(* PLC project Gaia V5.project, CODESYS CODESYS V3.5 SP22 Patch 2 *)
(* stored: creationDateTime 2026-10-19T15:55:08.3177105, modificationDateTime 2026-10-19T13:52:28.0800332 *)

TYPE DUT_EXC_DOSENSOR : STRUCT
  EXC_OUTPUT_SIGNAL : REAL;  (* [EXC : to other equipment] Dissolved oxygen measure *)
  UPI_INPUT_GLOBAL_LOCAL_FUXA : BOOL;  (* [UPI : functional units to equipment] From UPI_LOCAL_FUXA : global FUXA local active *)
  UPI_INPUT_GLOBAL_LOCAL_HMI : BOOL;  (* From UPI_LOCAL_HMI : global HMI local active *)
  UPI_INPUT_GLOBAL_LOCAL_WEBVISU : BOOL;  (* From UPI_LOCAL_webvisu : global HMI local active *)
END_STRUCT;
END_TYPE

TYPE DUT_IO_DOSENSOR : STRUCT
  INPUT_SIGNAL : DWORD;  (* [INPUT (field to PLC)] Analog input, raw value *)
  INPUT_SENSOR_FAULT : BOOL;  (* Digital input, sensor fault *)
  OUTPUT_CALIBRATION_HIGH : BOOL;  (* [OUTPUT (PLC to field)] Digital output, high calibration *)
  OUTPUT_CALIBRATION_LOW : BOOL;  (* Digital output, low calibration *)
END_STRUCT;
END_TYPE

TYPE DUT_INT_DOSENSOR : STRUCT
  FUXA_LOCAL_REQUEST : BOOL;  (* [Control mode] From FUXA : local request (pulse or maintained) *)
  FUXA_AUTO_REQUEST : BOOL;  (* From FUXA : auto request, releases the individual FUXA local *)
  HMI_LOCAL_REQUEST : BOOL;  (* From HMI : local request (pulse or maintained) *)
  HMI_AUTO_REQUEST : BOOL;  (* From HMI : auto request, releases the individual HMI local *)
  GLOBAL_LOCAL_FUXA : BOOL;  (* From UPI_LOCAL_FUXA : global FUXA local active *)
  GLOBAL_LOCAL_HMI : BOOL;  (* From UPI_LOCAL_HMI : global HMI local active *)
  LOCAL_FUXA_INDIVIDUAL : BOOL;  (* Memory : individual FUXA local, set by local request, reset by auto request *)
  LOCAL_HMI_INDIVIDUAL : BOOL;  (* Memory : individual HMI local, set by local request, reset by auto request *)
  LOCAL_HMI : BOOL;  (* Result : equipment in HMI local (individual or global), unless WEBVISU local is active *)
  LOCAL_FUXA : BOOL;  (* Result : equipment in FUXA local (individual or global), unless WEBVISU or HMI local is active *)
  WEBVISU_LOCAL_REQUEST : BOOL;  (* From WEBVISU : local request (pulse or maintained) *)
  WEBVISU_AUTO_REQUEST : BOOL;  (* From WEBVISU : auto request, releases the individual WEBVISU local *)
  LOCAL_WEBVISU_INDIVIDUAL : BOOL;  (* Memory : individual WEBVISU local, set by local request, reset by auto request *)
  LOCAL_WEBVISU : BOOL;  (* Result : equipment in WEBVISU local (individual or global), has priority *)
  AUTO : BOOL;  (* Result : no local mode, commands come from the functional units (UPI) *)
  SIGNAL_RAW : DWORD;  (* [Inputs] Raw analog input *)
  FAULT : BOOL;  (* Sensor fault (digital input) *)
  CALIB_HIGH_REQUEST : BOOL;  (* High calibration request from the active source *)
  CALIB_LOW_REQUEST : BOOL;  (* Low calibration request from the active source *)
  SIGNAL : REAL;  (* [Results] Scaled measure *)
  CALIB_HIGH : BOOL;  (* High calibration pulse to sensor (1 s) *)
  CALIB_LOW : BOOL;  (* Low calibration pulse to sensor (1 s) *)
  CALIB_DONE : BOOL;  (* Calibration done message (5 s) *)
  GLOBAL_LOCAL_WEBVISU : BOOL;  (* From UPI_LOCAL_WEBVISU : global local request *)
END_STRUCT;
END_TYPE

TYPE DUT_COM_DOSENSOR : STRUCT
  SCADA_INPUT_CALIBRATION_HIGH : BOOL;  (* [SCADA (FUXA) : input (to PLC)] Coil 1 | DO Calibration High *)
  SCADA_INPUT_CALIBRATION_LOW : BOOL;  (* Coil 2 | DO Calibration Low *)
  SCADA_INPUT_LOCAL_REQUEST : BOOL;  (* Coil 8 | DO Sensor Local Request *)
  SCADA_INPUT_AUTO_REQUEST : BOOL;  (* Coil 9 | DO Sensor Auto Request *)
  SCADA_OUTPUT_FAULT : BOOL;  (* [SCADA (FUXA) : output (from PLC)] DI 10001 | Do sensor fault *)
  SCADA_OUTPUT_CALIBRATION_DONE : BOOL;  (* DI 10002 | Do sensor calibration done *)
  SCADA_OUTPUT_LOCAL_FUXA_ACTIVE : BOOL;  (* DI 10013 | DO Sensor Local FUXA Active *)
  SCADA_OUTPUT_LOCAL_HMI_ACTIVE : BOOL;  (* DI 10014 | DO Sensor Local HMI Active *)
  SCADA_OUTPUT_SIGNAL : DUT_Union_Real_Word;  (* IR 89-90 | DO Sensor Signal *)
  HMI_INPUT_CALIBRATION_HIGH : BOOL;  (* [HMI (local panel, FUXA address + 1000) : input (to PLC)] Coil 1001 | DO Calibration High *)
  HMI_INPUT_CALIBRATION_LOW : BOOL;  (* Coil 1002 | DO Calibration Low *)
  HMI_INPUT_LOCAL_REQUEST : BOOL;  (* Coil 1008 | DO Sensor Local Request *)
  HMI_INPUT_AUTO_REQUEST : BOOL;  (* Coil 1009 | DO Sensor Auto Request *)
  HMI_OUTPUT_FAULT : BOOL;  (* [HMI (local panel, FUXA address + 1000) : output (from PLC)] DI 11001 | Do sensor fault *)
  HMI_OUTPUT_CALIBRATION_DONE : BOOL;  (* DI 11002 | Do sensor calibration done *)
  HMI_OUTPUT_LOCAL_ACTIVE : BOOL;  (* DI 11014 | DO Sensor Local Active *)
  HMI_OUTPUT_SIGNAL : DUT_Union_Real_Word;  (* IR 1089-1090 | DO Sensor Signal *)
  WEBVISU_INPUT_CALIBRATION_HIGH : BOOL;  (* DO Calibration High *)
  WEBVISU_INPUT_CALIBRATION_LOW : BOOL;  (* DO Calibration Low *)
  WEBVISU_INPUT_LOCAL_REQUEST : BOOL;  (* DO Sensor Local Request *)
  WEBVISU_INPUT_AUTO_REQUEST : BOOL;  (* DO Sensor Auto Request *)
  WEBVISU_OUTPUT_FAULT : BOOL;  (* Do sensor fault *)
  WEBVISU_OUTPUT_CALIBRATION_DONE : BOOL;  (* Do sensor calibration done *)
  WEBVISU_OUTPUT_LOCAL_ACTIVE : BOOL;  (* DO Sensor Local Active *)
  WEBVISU_OUTPUT_SIGNAL : DUT_Union_Real_Word;  (* DO Sensor Signal *)
  WEBVISU_OUTPUT_LOCAL_FUXA_ACTIVE : BOOL;  (* Effective FUXA local mode (masked by WEBVISU and HMI priority) *)
  WEBVISU_OUTPUT_LOCAL_HMI_ACTIVE : BOOL;  (* Effective HMI local mode (masked by WEBVISU priority) *)
END_STRUCT;
END_TYPE

TYPE DUT_INT_ADM100W : STRUCT
  FUXA_LOCAL_REQUEST : BOOL;  (* [Control mode] From FUXA : local request (pulse or maintained) *)
  FUXA_AUTO_REQUEST : BOOL;  (* From FUXA : auto request, releases the individual FUXA local *)
  HMI_LOCAL_REQUEST : BOOL;  (* From HMI : local request (pulse or maintained) *)
  HMI_AUTO_REQUEST : BOOL;  (* From HMI : auto request, releases the individual HMI local *)
  GLOBAL_LOCAL_FUXA : BOOL;  (* From UPI_LOCAL_FUXA : global FUXA local active *)
  GLOBAL_LOCAL_HMI : BOOL;  (* From UPI_LOCAL_HMI : global HMI local active *)
  LOCAL_FUXA_INDIVIDUAL : BOOL;  (* Memory : individual FUXA local, set by local request, reset by auto request *)
  LOCAL_HMI_INDIVIDUAL : BOOL;  (* Memory : individual HMI local, set by local request, reset by auto request *)
  LOCAL_HMI : BOOL;  (* Result : equipment in HMI local (individual or global), unless WEBVISU local is active *)
  LOCAL_FUXA : BOOL;  (* Result : equipment in FUXA local (individual or global), unless WEBVISU or HMI local is active *)
  AUTO : BOOL;  (* Result : no local mode, commands come from the functional units (UPI) *)
  ALARM_1 : BOOL;  (* [Alarms] Alarm 1 status *)
  ALARM_2 : BOOL;  (* Alarm 2 status *)
  ALARM_3 : BOOL;  (* Alarm 3 status *)
  ALARM_4 : BOOL;  (* Alarm 4 status *)
  ALARM_5 : BOOL;  (* Alarm 5 status *)
  ALARM_6 : BOOL;  (* Alarm 6 status *)
  ALARM_7 : BOOL;  (* Alarm 7 status *)
  ALARM_8 : BOOL;  (* Alarm 8 status *)
  ALARM_9 : BOOL;  (* Alarm 9 status *)
  ALARM_10 : BOOL;  (* Alarm 10 status *)
  FREQUENCY : REAL;  (* [Measures] Frequency | Hz *)
  L1_L2_VOLTAGE : REAL;  (* L1-L2 Voltage | V *)
  L1_N_VOLTAGE : REAL;  (* L1-N Voltage | V *)
  L1_CURRENT : REAL;  (* L1 Current | A *)
  L1_ACTIVE_POWER : REAL;  (* L1 Active Power | W *)
  L1_APPARENT_POWER : REAL;  (* L1 Apparent Power | VA *)
  L1_REACTIVE_POWER : REAL;  (* L1 Reactive Power | W *)
  L1_CURRENT_PHASE_ANGLE : REAL;  (* L1 Current Phase Angle | deg *)
  L1_POWER_FACTOR : REAL;  (* L1 Power Factor | - *)
  L1_VOLTAGE_THD : REAL;  (* L1 Voltage THD | % *)
  L1_CURRENT_THD : REAL;  (* L1 Current THD | % *)
  L1_MAX_LOAD : REAL;  (* L1 Max Load | % of 60 A *)
  L1_L2_VOLTAGE_PHASE_ANGLE : REAL;  (* L1-L2 Voltage Phase Angle | deg *)
  L2_L3_VOLTAGE : REAL;  (* L2-L3 Voltage | V *)
  L2_N_VOLTAGE : REAL;  (* L2-N Voltage | V *)
  L2_CURRENT : REAL;  (* L2 Current | A *)
  L2_ACTIVE_POWER : REAL;  (* L2 Active Power | W *)
  L2_APPARENT_POWER : REAL;  (* L2 Apparent Power | VA *)
  L2_REACTIVE_POWER : REAL;  (* L2 Reactive Power | W *)
  L2_CURRENT_PHASE_ANGLE : REAL;  (* L2 Current Phase Angle | deg *)
  L2_POWER_FACTOR : REAL;  (* L2 Power Factor | - *)
  L2_VOLTAGE_THD : REAL;  (* L2 Voltage THD | % *)
  L2_CURRENT_THD : REAL;  (* L2 Current THD | % *)
  L2_MAX_LOAD : REAL;  (* L2 Max Load | % of 60 A *)
  L1_L3_VOLTAGE_PHASE_ANGLE : REAL;  (* L1-L3 Voltage Phase Angle | deg *)
  L3_L1_VOLTAGE : REAL;  (* L3-L1 Voltage | V *)
  L3_N_VOLTAGE : REAL;  (* L3-N Voltage | V *)
  L3_CURRENT : REAL;  (* L3 Current | A *)
  L3_ACTIVE_POWER : REAL;  (* L3 Active Power | W *)
  L3_APPARENT_POWER : REAL;  (* L3 Apparent Power | VA *)
  L3_REACTIVE_POWER : REAL;  (* L3 Reactive Power | W *)
  L3_CURRENT_PHASE_ANGLE : REAL;  (* L3 Current Phase Angle | deg *)
  L3_POWER_FACTOR : REAL;  (* L3 Power Factor | - *)
  L3_VOLTAGE_THD : REAL;  (* L3 Voltage THD | % *)
  L3_CURRENT_THD : REAL;  (* L3 Current THD | % *)
  L3_MAX_LOAD : REAL;  (* L3 Max Load | % of 60 A *)
  INTERNAL_TEMPERATURE : REAL;  (* Internal Temperature | degC *)
  ACTIVE_ENERGY : REAL;  (* Active Energy | kWh *)
  APPARENT_ENERGY : REAL;  (* Apparent Energy | per ADM100W config *)
  REACTIVE_ENERGY : REAL;  (* Reactive Energy | kWh *)
  TOTAL_ACTIVE_POWER : REAL;  (* Total Active Power | W *)
  TOTAL_APPARENT_POWER : REAL;  (* Total Apparent Power | VA *)
  TOTAL_REACTIVE_POWER : REAL;  (* Total Reactive Power | W *)
  ALL_PHASE_POWER_FACTOR : REAL;  (* All Phase Power Factor | - *)
  WEBVISU_LOCAL_REQUEST : BOOL;  (* From WEBVISU : individual local request *)
  WEBVISU_AUTO_REQUEST : BOOL;  (* From WEBVISU : releases individual WEBVISU local (auto wins) *)
  GLOBAL_LOCAL_WEBVISU : BOOL;  (* From UPI_LOCAL_WEBVISU : global local request *)
  LOCAL_WEBVISU_INDIVIDUAL : BOOL;  (* Memory : individual WEBVISU local request *)
  LOCAL_WEBVISU : BOOL;  (* Effective WEBVISU local : highest source priority *)
END_STRUCT;
END_TYPE

TYPE DUT_COM_UPI_LOCAL_FUXA : STRUCT
  SCADA_INPUT_LOCAL_REQUEST : BOOL;  (* [SCADA (FUXA) : input (to PLC)] Coil 14 | Global Local FUXA Request *)
  SCADA_INPUT_AUTO_REQUEST : BOOL;  (* Coil 15 | Global Auto FUXA Request *)
  SCADA_OUTPUT_LOCAL_ACTIVE : BOOL;  (* [SCADA (FUXA) : output (from PLC)] DI 10019 | Global Local FUXA Active *)
END_STRUCT;
END_TYPE

TYPE DUT_IO_ADM100W : STRUCT
  SPARE : BOOL;  (* Placeholder, structure not used yet *)
END_STRUCT;
END_TYPE

TYPE DUT_COM_ADM100W : STRUCT
  COM_INPUT_IR : ARRAY[0..87] OF WORD;  (* [COM : Modbus RTU, input (equipment to PLC)] Input registers 0..87, 32-bit float, MSW first (ABCD) *)
  COM_INPUT_COILS : ARRAY[0..1] OF BYTE;  (* Coils 0..9 = alarms 1..10 (byte.bit) *)
  SCADA_INPUT_LOCAL_REQUEST : BOOL;  (* [SCADA (FUXA) : input (to PLC)] Coil 12 | ADM100W Local Request *)
  SCADA_INPUT_AUTO_REQUEST : BOOL;  (* Coil 13 | ADM100W Auto Request *)
  SCADA_OUTPUT_ALARM_1_STATUS : BOOL;  (* [SCADA (FUXA) : output (from PLC)] DI 10003 | ADM100W Alarm 1 Status *)
  SCADA_OUTPUT_ALARM_2_STATUS : BOOL;  (* DI 10004 | ADM100W Alarm 2 Status *)
  SCADA_OUTPUT_ALARM_3_STATUS : BOOL;  (* DI 10005 | ADM100W Alarm 3 Status *)
  SCADA_OUTPUT_ALARM_4_STATUS : BOOL;  (* DI 10006 | ADM100W Alarm 4 Status *)
  SCADA_OUTPUT_ALARM_5_STATUS : BOOL;  (* DI 10007 | ADM100W Alarm 5 Status *)
  SCADA_OUTPUT_ALARM_6_STATUS : BOOL;  (* DI 10008 | ADM100W Alarm 6 Status *)
  SCADA_OUTPUT_ALARM_7_STATUS : BOOL;  (* DI 10009 | ADM100W Alarm 7 Status *)
  SCADA_OUTPUT_ALARM_8_STATUS : BOOL;  (* DI 10010 | ADM100W Alarm 8 Status *)
  SCADA_OUTPUT_ALARM_9_STATUS : BOOL;  (* DI 10011 | ADM100W Alarm 9 Status *)
  SCADA_OUTPUT_ALARM_10_STATUS : BOOL;  (* DI 10012 | ADM100W Alarm 10 Status *)
  SCADA_OUTPUT_LOCAL_FUXA_ACTIVE : BOOL;  (* DI 10017 | ADM100W Local FUXA Active *)
  SCADA_OUTPUT_LOCAL_HMI_ACTIVE : BOOL;  (* DI 10018 | ADM100W Local HMI Active *)
  SCADA_OUTPUT_FREQUENCY : DUT_Union_Real_Word;  (* IR 1-2 | ADM100W Frequency | Hz *)
  SCADA_OUTPUT_L1_L2_VOLTAGE : DUT_Union_Real_Word;  (* IR 3-4 | ADM100W L1-L2 Voltage | V *)
  SCADA_OUTPUT_L1_N_VOLTAGE : DUT_Union_Real_Word;  (* IR 5-6 | ADM100W L1-N Voltage | V *)
  SCADA_OUTPUT_L1_CURRENT : DUT_Union_Real_Word;  (* IR 7-8 | ADM100W L1 Current | A *)
  SCADA_OUTPUT_L1_ACTIVE_POWER : DUT_Union_Real_Word;  (* IR 9-10 | ADM100W L1 Active Power *)
  SCADA_OUTPUT_L1_APPARENT_POWER : DUT_Union_Real_Word;  (* IR 11-12 | ADM100W L1 Apparent Power *)
  SCADA_OUTPUT_L1_REACTIVE_POWER : DUT_Union_Real_Word;  (* IR 13-14 | ADM100W L1 Reactive Power *)
  SCADA_OUTPUT_L1_CURRENT_PHASE_ANGLE : DUT_Union_Real_Word;  (* IR 15-16 | ADM100W L1 Current Phase Angle | deg *)
  SCADA_OUTPUT_L1_POWER_FACTOR : DUT_Union_Real_Word;  (* IR 17-18 | ADM100W L1 Power Factor *)
  SCADA_OUTPUT_L1_VOLTAGE_THD : DUT_Union_Real_Word;  (* IR 19-20 | ADM100W L1 Voltage THD | % *)
  SCADA_OUTPUT_L1_CURRENT_THD : DUT_Union_Real_Word;  (* IR 21-22 | ADM100W L1 Current THD | % *)
  SCADA_OUTPUT_L1_MAX_LOAD : DUT_Union_Real_Word;  (* IR 23-24 | ADM100W L1 Max Load *)
  SCADA_OUTPUT_L1_L2_VOLTAGE_PHASE_ANGLE : DUT_Union_Real_Word;  (* IR 25-26 | ADM100W L1-L2 Voltage Phase Angle | deg *)
  SCADA_OUTPUT_L2_L3_VOLTAGE : DUT_Union_Real_Word;  (* IR 27-28 | ADM100W L2-L3 Voltage | V *)
  SCADA_OUTPUT_L2_N_VOLTAGE : DUT_Union_Real_Word;  (* IR 29-30 | ADM100W L2-N Voltage | V *)
  SCADA_OUTPUT_L2_CURRENT : DUT_Union_Real_Word;  (* IR 31-32 | ADM100W L2 Current | A *)
  SCADA_OUTPUT_L2_ACTIVE_POWER : DUT_Union_Real_Word;  (* IR 33-34 | ADM100W L2 Active Power *)
  SCADA_OUTPUT_L2_APPARENT_POWER : DUT_Union_Real_Word;  (* IR 35-36 | ADM100W L2 Apparent Power *)
  SCADA_OUTPUT_L2_REACTIVE_POWER : DUT_Union_Real_Word;  (* IR 37-38 | ADM100W L2 Reactive Power *)
  SCADA_OUTPUT_L2_CURRENT_PHASE_ANGLE : DUT_Union_Real_Word;  (* IR 39-40 | ADM100W L2 Current Phase Angle | deg *)
  SCADA_OUTPUT_L2_POWER_FACTOR : DUT_Union_Real_Word;  (* IR 41-42 | ADM100W L2 Power Factor *)
  SCADA_OUTPUT_L2_VOLTAGE_THD : DUT_Union_Real_Word;  (* IR 43-44 | ADM100W L2 Voltage THD | % *)
  SCADA_OUTPUT_L2_CURRENT_THD : DUT_Union_Real_Word;  (* IR 45-46 | ADM100W L2 Current THD | % *)
  SCADA_OUTPUT_L2_MAX_LOAD : DUT_Union_Real_Word;  (* IR 47-48 | ADM100W L2 Max Load *)
  SCADA_OUTPUT_L1_L3_VOLTAGE_PHASE_ANGLE : DUT_Union_Real_Word;  (* IR 49-50 | ADM100W L1-L3 Voltage Phase Angle | deg *)
  SCADA_OUTPUT_L3_L1_VOLTAGE : DUT_Union_Real_Word;  (* IR 51-52 | ADM100W L3-L1 Voltage | V *)
  SCADA_OUTPUT_L3_N_VOLTAGE : DUT_Union_Real_Word;  (* IR 53-54 | ADM100W L3-N Voltage | V *)
  SCADA_OUTPUT_L3_CURRENT : DUT_Union_Real_Word;  (* IR 55-56 | ADM100W L3 Current | A *)
  SCADA_OUTPUT_L3_ACTIVE_POWER : DUT_Union_Real_Word;  (* IR 57-58 | ADM100W L3 Active Power *)
  SCADA_OUTPUT_L3_APPARENT_POWER : DUT_Union_Real_Word;  (* IR 59-60 | ADM100W L3 Apparent Power *)
  SCADA_OUTPUT_L3_REACTIVE_POWER : DUT_Union_Real_Word;  (* IR 61-62 | ADM100W L3 Reactive Power *)
  SCADA_OUTPUT_L3_CURRENT_PHASE_ANGLE : DUT_Union_Real_Word;  (* IR 63-64 | ADM100W L3 Current Phase Angle | deg *)
  SCADA_OUTPUT_L3_POWER_FACTOR : DUT_Union_Real_Word;  (* IR 65-66 | ADM100W L3 Power Factor *)
  SCADA_OUTPUT_L3_VOLTAGE_THD : DUT_Union_Real_Word;  (* IR 67-68 | ADM100W L3 Voltage THD | % *)
  SCADA_OUTPUT_L3_CURRENT_THD : DUT_Union_Real_Word;  (* IR 69-70 | ADM100W L3 Current THD | % *)
  SCADA_OUTPUT_L3_MAX_LOAD : DUT_Union_Real_Word;  (* IR 71-72 | ADM100W L3 Max Load *)
  SCADA_OUTPUT_INTERNAL_TEMPERATURE : DUT_Union_Real_Word;  (* IR 73-74 | ADM100W Internal Temperature *)
  SCADA_OUTPUT_ACTIVE_ENERGY : DUT_Union_Real_Word;  (* IR 75-76 | ADM100W Active Energy *)
  SCADA_OUTPUT_APPARENT_ENERGY : DUT_Union_Real_Word;  (* IR 77-78 | ADM100W Apparent Energy *)
  SCADA_OUTPUT_REACTIVE_ENERGY : DUT_Union_Real_Word;  (* IR 79-80 | ADM100W Reactive Energy *)
  SCADA_OUTPUT_TOTAL_ACTIVE_POWER : DUT_Union_Real_Word;  (* IR 81-82 | ADM100W Total Active Power *)
  SCADA_OUTPUT_TOTAL_APPARENT_POWER : DUT_Union_Real_Word;  (* IR 83-84 | ADM100W Total Apparent Power *)
  SCADA_OUTPUT_TOTAL_REACTIVE_POWER : DUT_Union_Real_Word;  (* IR 85-86 | ADM100W Total Reactive Power *)
  SCADA_OUTPUT_ALL_PHASE_POWER_FACTOR : DUT_Union_Real_Word;  (* IR 87-88 | ADM100W All Phase Power Factor *)
  HMI_INPUT_LOCAL_REQUEST : BOOL;  (* [HMI (local panel, FUXA address + 1000) : input (to PLC)] Coil 1012 | ADM100W Local Request *)
  HMI_INPUT_AUTO_REQUEST : BOOL;  (* Coil 1013 | ADM100W Auto Request *)
  HMI_OUTPUT_ALARM_1_STATUS : BOOL;  (* [HMI (local panel, FUXA address + 1000) : output (from PLC)] DI 11003 | ADM100W Alarm 1 Status *)
  HMI_OUTPUT_ALARM_2_STATUS : BOOL;  (* DI 11004 | ADM100W Alarm 2 Status *)
  HMI_OUTPUT_ALARM_3_STATUS : BOOL;  (* DI 11005 | ADM100W Alarm 3 Status *)
  HMI_OUTPUT_ALARM_4_STATUS : BOOL;  (* DI 11006 | ADM100W Alarm 4 Status *)
  HMI_OUTPUT_ALARM_5_STATUS : BOOL;  (* DI 11007 | ADM100W Alarm 5 Status *)
  HMI_OUTPUT_ALARM_6_STATUS : BOOL;  (* DI 11008 | ADM100W Alarm 6 Status *)
  HMI_OUTPUT_ALARM_7_STATUS : BOOL;  (* DI 11009 | ADM100W Alarm 7 Status *)
  HMI_OUTPUT_ALARM_8_STATUS : BOOL;  (* DI 11010 | ADM100W Alarm 8 Status *)
  HMI_OUTPUT_ALARM_9_STATUS : BOOL;  (* DI 11011 | ADM100W Alarm 9 Status *)
  HMI_OUTPUT_ALARM_10_STATUS : BOOL;  (* DI 11012 | ADM100W Alarm 10 Status *)
  HMI_OUTPUT_LOCAL_ACTIVE : BOOL;  (* DI 11018 | ADM100W Local Active *)
  HMI_OUTPUT_FREQUENCY : DUT_Union_Real_Word;  (* IR 1001-1002 | ADM100W Frequency | Hz *)
  HMI_OUTPUT_L1_L2_VOLTAGE : DUT_Union_Real_Word;  (* IR 1003-1004 | ADM100W L1-L2 Voltage | V *)
  HMI_OUTPUT_L1_N_VOLTAGE : DUT_Union_Real_Word;  (* IR 1005-1006 | ADM100W L1-N Voltage | V *)
  HMI_OUTPUT_L1_CURRENT : DUT_Union_Real_Word;  (* IR 1007-1008 | ADM100W L1 Current | A *)
  HMI_OUTPUT_L1_ACTIVE_POWER : DUT_Union_Real_Word;  (* IR 1009-1010 | ADM100W L1 Active Power *)
  HMI_OUTPUT_L1_APPARENT_POWER : DUT_Union_Real_Word;  (* IR 1011-1012 | ADM100W L1 Apparent Power *)
  HMI_OUTPUT_L1_REACTIVE_POWER : DUT_Union_Real_Word;  (* IR 1013-1014 | ADM100W L1 Reactive Power *)
  HMI_OUTPUT_L1_CURRENT_PHASE_ANGLE : DUT_Union_Real_Word;  (* IR 1015-1016 | ADM100W L1 Current Phase Angle | deg *)
  HMI_OUTPUT_L1_POWER_FACTOR : DUT_Union_Real_Word;  (* IR 1017-1018 | ADM100W L1 Power Factor *)
  HMI_OUTPUT_L1_VOLTAGE_THD : DUT_Union_Real_Word;  (* IR 1019-1020 | ADM100W L1 Voltage THD | % *)
  HMI_OUTPUT_L1_CURRENT_THD : DUT_Union_Real_Word;  (* IR 1021-1022 | ADM100W L1 Current THD | % *)
  HMI_OUTPUT_L1_MAX_LOAD : DUT_Union_Real_Word;  (* IR 1023-1024 | ADM100W L1 Max Load *)
  HMI_OUTPUT_L1_L2_VOLTAGE_PHASE_ANGLE : DUT_Union_Real_Word;  (* IR 1025-1026 | ADM100W L1-L2 Voltage Phase Angle | deg *)
  HMI_OUTPUT_L2_L3_VOLTAGE : DUT_Union_Real_Word;  (* IR 1027-1028 | ADM100W L2-L3 Voltage | V *)
  HMI_OUTPUT_L2_N_VOLTAGE : DUT_Union_Real_Word;  (* IR 1029-1030 | ADM100W L2-N Voltage | V *)
  HMI_OUTPUT_L2_CURRENT : DUT_Union_Real_Word;  (* IR 1031-1032 | ADM100W L2 Current | A *)
  HMI_OUTPUT_L2_ACTIVE_POWER : DUT_Union_Real_Word;  (* IR 1033-1034 | ADM100W L2 Active Power *)
  HMI_OUTPUT_L2_APPARENT_POWER : DUT_Union_Real_Word;  (* IR 1035-1036 | ADM100W L2 Apparent Power *)
  HMI_OUTPUT_L2_REACTIVE_POWER : DUT_Union_Real_Word;  (* IR 1037-1038 | ADM100W L2 Reactive Power *)
  HMI_OUTPUT_L2_CURRENT_PHASE_ANGLE : DUT_Union_Real_Word;  (* IR 1039-1040 | ADM100W L2 Current Phase Angle | deg *)
  HMI_OUTPUT_L2_POWER_FACTOR : DUT_Union_Real_Word;  (* IR 1041-1042 | ADM100W L2 Power Factor *)
  HMI_OUTPUT_L2_VOLTAGE_THD : DUT_Union_Real_Word;  (* IR 1043-1044 | ADM100W L2 Voltage THD | % *)
  HMI_OUTPUT_L2_CURRENT_THD : DUT_Union_Real_Word;  (* IR 1045-1046 | ADM100W L2 Current THD | % *)
  HMI_OUTPUT_L2_MAX_LOAD : DUT_Union_Real_Word;  (* IR 1047-1048 | ADM100W L2 Max Load *)
  HMI_OUTPUT_L1_L3_VOLTAGE_PHASE_ANGLE : DUT_Union_Real_Word;  (* IR 1049-1050 | ADM100W L1-L3 Voltage Phase Angle | deg *)
  HMI_OUTPUT_L3_L1_VOLTAGE : DUT_Union_Real_Word;  (* IR 1051-1052 | ADM100W L3-L1 Voltage | V *)
  HMI_OUTPUT_L3_N_VOLTAGE : DUT_Union_Real_Word;  (* IR 1053-1054 | ADM100W L3-N Voltage | V *)
  HMI_OUTPUT_L3_CURRENT : DUT_Union_Real_Word;  (* IR 1055-1056 | ADM100W L3 Current | A *)
  HMI_OUTPUT_L3_ACTIVE_POWER : DUT_Union_Real_Word;  (* IR 1057-1058 | ADM100W L3 Active Power *)
  HMI_OUTPUT_L3_APPARENT_POWER : DUT_Union_Real_Word;  (* IR 1059-1060 | ADM100W L3 Apparent Power *)
  HMI_OUTPUT_L3_REACTIVE_POWER : DUT_Union_Real_Word;  (* IR 1061-1062 | ADM100W L3 Reactive Power *)
  HMI_OUTPUT_L3_CURRENT_PHASE_ANGLE : DUT_Union_Real_Word;  (* IR 1063-1064 | ADM100W L3 Current Phase Angle | deg *)
  HMI_OUTPUT_L3_POWER_FACTOR : DUT_Union_Real_Word;  (* IR 1065-1066 | ADM100W L3 Power Factor *)
  HMI_OUTPUT_L3_VOLTAGE_THD : DUT_Union_Real_Word;  (* IR 1067-1068 | ADM100W L3 Voltage THD | % *)
  HMI_OUTPUT_L3_CURRENT_THD : DUT_Union_Real_Word;  (* IR 1069-1070 | ADM100W L3 Current THD | % *)
  HMI_OUTPUT_L3_MAX_LOAD : DUT_Union_Real_Word;  (* IR 1071-1072 | ADM100W L3 Max Load *)
  HMI_OUTPUT_INTERNAL_TEMPERATURE : DUT_Union_Real_Word;  (* IR 1073-1074 | ADM100W Internal Temperature *)
  HMI_OUTPUT_ACTIVE_ENERGY : DUT_Union_Real_Word;  (* IR 1075-1076 | ADM100W Active Energy *)
  HMI_OUTPUT_APPARENT_ENERGY : DUT_Union_Real_Word;  (* IR 1077-1078 | ADM100W Apparent Energy *)
  HMI_OUTPUT_REACTIVE_ENERGY : DUT_Union_Real_Word;  (* IR 1079-1080 | ADM100W Reactive Energy *)
  HMI_OUTPUT_TOTAL_ACTIVE_POWER : DUT_Union_Real_Word;  (* IR 1081-1082 | ADM100W Total Active Power *)
  HMI_OUTPUT_TOTAL_APPARENT_POWER : DUT_Union_Real_Word;  (* IR 1083-1084 | ADM100W Total Apparent Power *)
  HMI_OUTPUT_TOTAL_REACTIVE_POWER : DUT_Union_Real_Word;  (* IR 1085-1086 | ADM100W Total Reactive Power *)
  HMI_OUTPUT_ALL_PHASE_POWER_FACTOR : DUT_Union_Real_Word;  (* IR 1087-1088 | ADM100W All Phase Power Factor *)
  WEBVISU_INPUT_LOCAL_REQUEST : BOOL;  (* [WEBVISU : direct IEC variable] ADM100W Local Request *)
  WEBVISU_INPUT_AUTO_REQUEST : BOOL;  (* [WEBVISU : direct IEC variable] ADM100W Auto Request *)
  WEBVISU_OUTPUT_ALARM_1_STATUS : BOOL;  (* [WEBVISU : direct IEC variable] ADM100W Alarm 1 Status *)
  WEBVISU_OUTPUT_ALARM_2_STATUS : BOOL;  (* [WEBVISU : direct IEC variable] ADM100W Alarm 2 Status *)
  WEBVISU_OUTPUT_ALARM_3_STATUS : BOOL;  (* [WEBVISU : direct IEC variable] ADM100W Alarm 3 Status *)
  WEBVISU_OUTPUT_ALARM_4_STATUS : BOOL;  (* [WEBVISU : direct IEC variable] ADM100W Alarm 4 Status *)
  WEBVISU_OUTPUT_ALARM_5_STATUS : BOOL;  (* [WEBVISU : direct IEC variable] ADM100W Alarm 5 Status *)
  WEBVISU_OUTPUT_ALARM_6_STATUS : BOOL;  (* [WEBVISU : direct IEC variable] ADM100W Alarm 6 Status *)
  WEBVISU_OUTPUT_ALARM_7_STATUS : BOOL;  (* [WEBVISU : direct IEC variable] ADM100W Alarm 7 Status *)
  WEBVISU_OUTPUT_ALARM_8_STATUS : BOOL;  (* [WEBVISU : direct IEC variable] ADM100W Alarm 8 Status *)
  WEBVISU_OUTPUT_ALARM_9_STATUS : BOOL;  (* [WEBVISU : direct IEC variable] ADM100W Alarm 9 Status *)
  WEBVISU_OUTPUT_ALARM_10_STATUS : BOOL;  (* [WEBVISU : direct IEC variable] ADM100W Alarm 10 Status *)
  WEBVISU_OUTPUT_LOCAL_ACTIVE : BOOL;  (* [WEBVISU : direct IEC variable] ADM100W Local Active *)
  WEBVISU_OUTPUT_FREQUENCY : DUT_Union_Real_Word;  (* [WEBVISU : direct IEC variable] ADM100W Frequency | Hz *)
  WEBVISU_OUTPUT_L1_L2_VOLTAGE : DUT_Union_Real_Word;  (* [WEBVISU : direct IEC variable] ADM100W L1-L2 Voltage | V *)
  WEBVISU_OUTPUT_L1_N_VOLTAGE : DUT_Union_Real_Word;  (* [WEBVISU : direct IEC variable] ADM100W L1-N Voltage | V *)
  WEBVISU_OUTPUT_L1_CURRENT : DUT_Union_Real_Word;  (* [WEBVISU : direct IEC variable] ADM100W L1 Current | A *)
  WEBVISU_OUTPUT_L1_ACTIVE_POWER : DUT_Union_Real_Word;  (* [WEBVISU : direct IEC variable] ADM100W L1 Active Power *)
  WEBVISU_OUTPUT_L1_APPARENT_POWER : DUT_Union_Real_Word;  (* [WEBVISU : direct IEC variable] ADM100W L1 Apparent Power *)
  WEBVISU_OUTPUT_L1_REACTIVE_POWER : DUT_Union_Real_Word;  (* [WEBVISU : direct IEC variable] ADM100W L1 Reactive Power *)
  WEBVISU_OUTPUT_L1_CURRENT_PHASE_ANGLE : DUT_Union_Real_Word;  (* [WEBVISU : direct IEC variable] ADM100W L1 Current Phase Angle | deg *)
  WEBVISU_OUTPUT_L1_POWER_FACTOR : DUT_Union_Real_Word;  (* [WEBVISU : direct IEC variable] ADM100W L1 Power Factor *)
  WEBVISU_OUTPUT_L1_VOLTAGE_THD : DUT_Union_Real_Word;  (* [WEBVISU : direct IEC variable] ADM100W L1 Voltage THD | % *)
  WEBVISU_OUTPUT_L1_CURRENT_THD : DUT_Union_Real_Word;  (* [WEBVISU : direct IEC variable] ADM100W L1 Current THD | % *)
  WEBVISU_OUTPUT_L1_MAX_LOAD : DUT_Union_Real_Word;  (* [WEBVISU : direct IEC variable] ADM100W L1 Max Load *)
  WEBVISU_OUTPUT_L1_L2_VOLTAGE_PHASE_ANGLE : DUT_Union_Real_Word;  (* [WEBVISU : direct IEC variable] ADM100W L1-L2 Voltage Phase Angle | deg *)
  WEBVISU_OUTPUT_L2_L3_VOLTAGE : DUT_Union_Real_Word;  (* [WEBVISU : direct IEC variable] ADM100W L2-L3 Voltage | V *)
  WEBVISU_OUTPUT_L2_N_VOLTAGE : DUT_Union_Real_Word;  (* [WEBVISU : direct IEC variable] ADM100W L2-N Voltage | V *)
  WEBVISU_OUTPUT_L2_CURRENT : DUT_Union_Real_Word;  (* [WEBVISU : direct IEC variable] ADM100W L2 Current | A *)
  WEBVISU_OUTPUT_L2_ACTIVE_POWER : DUT_Union_Real_Word;  (* [WEBVISU : direct IEC variable] ADM100W L2 Active Power *)
  WEBVISU_OUTPUT_L2_APPARENT_POWER : DUT_Union_Real_Word;  (* [WEBVISU : direct IEC variable] ADM100W L2 Apparent Power *)
  WEBVISU_OUTPUT_L2_REACTIVE_POWER : DUT_Union_Real_Word;  (* [WEBVISU : direct IEC variable] ADM100W L2 Reactive Power *)
  WEBVISU_OUTPUT_L2_CURRENT_PHASE_ANGLE : DUT_Union_Real_Word;  (* [WEBVISU : direct IEC variable] ADM100W L2 Current Phase Angle | deg *)
  WEBVISU_OUTPUT_L2_POWER_FACTOR : DUT_Union_Real_Word;  (* [WEBVISU : direct IEC variable] ADM100W L2 Power Factor *)
  WEBVISU_OUTPUT_L2_VOLTAGE_THD : DUT_Union_Real_Word;  (* [WEBVISU : direct IEC variable] ADM100W L2 Voltage THD | % *)
  WEBVISU_OUTPUT_L2_CURRENT_THD : DUT_Union_Real_Word;  (* [WEBVISU : direct IEC variable] ADM100W L2 Current THD | % *)
  WEBVISU_OUTPUT_L2_MAX_LOAD : DUT_Union_Real_Word;  (* [WEBVISU : direct IEC variable] ADM100W L2 Max Load *)
  WEBVISU_OUTPUT_L1_L3_VOLTAGE_PHASE_ANGLE : DUT_Union_Real_Word;  (* [WEBVISU : direct IEC variable] ADM100W L1-L3 Voltage Phase Angle | deg *)
  WEBVISU_OUTPUT_L3_L1_VOLTAGE : DUT_Union_Real_Word;  (* [WEBVISU : direct IEC variable] ADM100W L3-L1 Voltage | V *)
  WEBVISU_OUTPUT_L3_N_VOLTAGE : DUT_Union_Real_Word;  (* [WEBVISU : direct IEC variable] ADM100W L3-N Voltage | V *)
  WEBVISU_OUTPUT_L3_CURRENT : DUT_Union_Real_Word;  (* [WEBVISU : direct IEC variable] ADM100W L3 Current | A *)
  WEBVISU_OUTPUT_L3_ACTIVE_POWER : DUT_Union_Real_Word;  (* [WEBVISU : direct IEC variable] ADM100W L3 Active Power *)
  WEBVISU_OUTPUT_L3_APPARENT_POWER : DUT_Union_Real_Word;  (* [WEBVISU : direct IEC variable] ADM100W L3 Apparent Power *)
  WEBVISU_OUTPUT_L3_REACTIVE_POWER : DUT_Union_Real_Word;  (* [WEBVISU : direct IEC variable] ADM100W L3 Reactive Power *)
  WEBVISU_OUTPUT_L3_CURRENT_PHASE_ANGLE : DUT_Union_Real_Word;  (* [WEBVISU : direct IEC variable] ADM100W L3 Current Phase Angle | deg *)
  WEBVISU_OUTPUT_L3_POWER_FACTOR : DUT_Union_Real_Word;  (* [WEBVISU : direct IEC variable] ADM100W L3 Power Factor *)
  WEBVISU_OUTPUT_L3_VOLTAGE_THD : DUT_Union_Real_Word;  (* [WEBVISU : direct IEC variable] ADM100W L3 Voltage THD | % *)
  WEBVISU_OUTPUT_L3_CURRENT_THD : DUT_Union_Real_Word;  (* [WEBVISU : direct IEC variable] ADM100W L3 Current THD | % *)
  WEBVISU_OUTPUT_L3_MAX_LOAD : DUT_Union_Real_Word;  (* [WEBVISU : direct IEC variable] ADM100W L3 Max Load *)
  WEBVISU_OUTPUT_INTERNAL_TEMPERATURE : DUT_Union_Real_Word;  (* [WEBVISU : direct IEC variable] ADM100W Internal Temperature *)
  WEBVISU_OUTPUT_ACTIVE_ENERGY : DUT_Union_Real_Word;  (* [WEBVISU : direct IEC variable] ADM100W Active Energy *)
  WEBVISU_OUTPUT_APPARENT_ENERGY : DUT_Union_Real_Word;  (* [WEBVISU : direct IEC variable] ADM100W Apparent Energy *)
  WEBVISU_OUTPUT_REACTIVE_ENERGY : DUT_Union_Real_Word;  (* [WEBVISU : direct IEC variable] ADM100W Reactive Energy *)
  WEBVISU_OUTPUT_TOTAL_ACTIVE_POWER : DUT_Union_Real_Word;  (* [WEBVISU : direct IEC variable] ADM100W Total Active Power *)
  WEBVISU_OUTPUT_TOTAL_APPARENT_POWER : DUT_Union_Real_Word;  (* [WEBVISU : direct IEC variable] ADM100W Total Apparent Power *)
  WEBVISU_OUTPUT_TOTAL_REACTIVE_POWER : DUT_Union_Real_Word;  (* [WEBVISU : direct IEC variable] ADM100W Total Reactive Power *)
  WEBVISU_OUTPUT_ALL_PHASE_POWER_FACTOR : DUT_Union_Real_Word;  (* [WEBVISU : direct IEC variable] ADM100W All Phase Power Factor *)
  WEBVISU_OUTPUT_LOCAL_FUXA_ACTIVE : BOOL;  (* Effective FUXA local mode (masked by WEBVISU and HMI priority) *)
  WEBVISU_OUTPUT_LOCAL_HMI_ACTIVE : BOOL;  (* Effective HMI local mode (masked by WEBVISU priority) *)
END_STRUCT;
END_TYPE

TYPE DUT_EXC_ADM100W : STRUCT
  EXC_OUTPUT_FREQUENCY : REAL;  (* [EXC : to other equipment] Hz *)
  EXC_OUTPUT_L1_N_VOLTAGE : REAL;  (* V *)
  EXC_OUTPUT_L1_CURRENT : REAL;  (* A *)
  EXC_OUTPUT_L1_ACTIVE_POWER : REAL;  (* W *)
  EXC_OUTPUT_L1_APPARENT_POWER : REAL;  (* VA *)
  EXC_OUTPUT_L1_REACTIVE_POWER : REAL;  (* VAr *)
  EXC_OUTPUT_L1_POWER_FACTOR : REAL;  (* - *)
  EXC_OUTPUT_L1_VOLTAGE_THD : REAL;  (* % *)
  EXC_OUTPUT_L1_CURRENT_THD : REAL;  (* % *)
  EXC_OUTPUT_L1_MAX_LOAD : REAL;  (* % of 60 A *)
  EXC_OUTPUT_INTERNAL_TEMPERATURE : REAL;  (* degC *)
  EXC_OUTPUT_ACTIVE_ENERGY : REAL;  (* kWh *)
  EXC_OUTPUT_DATA_VALID : BOOL;  (* FALSE = values not usable. Not managed yet (no Modbus diagnostic) *)
  UPI_INPUT_GLOBAL_LOCAL_FUXA : BOOL;  (* [UPI : functional units to equipment] From UPI_LOCAL_FUXA : global FUXA local active *)
  UPI_INPUT_GLOBAL_LOCAL_HMI : BOOL;  (* From UPI_LOCAL_HMI : global HMI local active *)
  UPI_INPUT_GLOBAL_LOCAL_WEBVISU : BOOL;  (* From UPI_LOCAL_WEBVISU : global WEBVISU local active *)
END_STRUCT;
END_TYPE

TYPE DUT_COM_DIP1500 : STRUCT
  COM_INPUT_IR : ARRAY[0..4] OF WORD;  (* [COM : Modbus RTU, input (equipment to PLC)] Input registers 0x3001..0x3005 *)
  COM_INPUT_HR_COUNTERS : ARRAY[0..3] OF WORD;  (* Holding registers 0x4007..0x400A (read) *)
  COM_OUTPUT_COILS : ARRAY[0..3] OF BOOL;  (* [COM : Modbus RTU, output (PLC to equipment)] Coils 0x0001..0x0004 *)
  COM_OUTPUT_HR_CMD : ARRAY[0..5] OF WORD;  (* Holding registers 0x4001..0x4006 (write) *)
  COM_OUTPUT_HR_CONFIG : ARRAY[0..6] OF WORD;  (* Holding registers 0x400B..0x4011 (write) *)
  COM_OUTPUT_CMD_TRIGGER : BOOL;  (* Rising edge trigger of the command write channel(s), mapped in the Modbus slave I/O mapping *)
  COM_OUTPUT_CONFIG_TRIGGER : BOOL;  (* Rising edge trigger of the configuration write channel, mapped in the Modbus slave I/O mapping *)
  SCADA_INPUT_MOTOR_START_STOP : BOOL;  (* [SCADA (FUXA) : input (to PLC)] Coil 3 | DIP1500 Motor Start Stop *)
  SCADA_INPUT_MOTOR_DIRECTION : BOOL;  (* Coil 4 | DIP1500 Motor Direction *)
  SCADA_INPUT_FLASH_SAVE : BOOL;  (* Coil 5 | DIP1500 Flash Save *)
  SCADA_INPUT_OPERATION_MODE : BOOL;  (* Coil 6 | DIP1500 Operation Mode *)
  SCADA_INPUT_PARAM_WRITE_ENABLE : BOOL;  (* Coil 7 | DIP1500 Parameter Write Enable *)
  SCADA_INPUT_LOCAL_REQUEST : BOOL;  (* Coil 10 | DIP1500 Local Request *)
  SCADA_INPUT_AUTO_REQUEST : BOOL;  (* Coil 11 | DIP1500 Auto Request *)
  SCADA_INPUT_FOOT_SWITCH_INPUT_MODE : WORD;  (* HR 9 | DIP1500 Foot Switch Input Mode *)
  SCADA_INPUT_LIQUID_LEVEL_INPUT_MODE : WORD;  (* HR 10 | DIP1500 Liquid Level Input Mode *)
  SCADA_INPUT_STATE_OUTPUT_MODE : WORD;  (* HR 11 | DIP1500 State Output Mode *)
  SCADA_INPUT_COMMUNICATION_ADDRESS : WORD;  (* HR 12 | DIP1500 Communication Address *)
  SCADA_INPUT_BAUD_RATE_INDEX : WORD;  (* HR 13 | DIP1500 Baud Rate Index | index *)
  SCADA_INPUT_MOTOR_SPEED : DUT_Union_Real_Word;  (* HR 1-2 | DIP1500 Motor Speed | rpm *)
  SCADA_INPUT_MAX_MOTOR_SPEED : DUT_Union_Real_Word;  (* HR 3-4 | DIP1500 Max Motor Speed | rpm *)
  SCADA_INPUT_RUN_TIME_OR_VOLUME_SETPOINT : DUT_Union_Real_Word;  (* HR 5-6 | DIP1500 Run Time Or Volume Setpoint | ms (time mode) / ml (volume mode) *)
  SCADA_INPUT_FLOW_RATE_OR_SPEED_CALIBRATION_COEFFICIENT : DUT_Union_Real_Word;  (* HR 7-8 | DIP1500 Flow Rate Or Speed Calibration Coefficient | ml/min or rpm *)
  SCADA_OUTPUT_LOCAL_FUXA_ACTIVE : BOOL;  (* [SCADA (FUXA) : output (from PLC)] DI 10015 | DIP1500 Local FUXA Active *)
  SCADA_OUTPUT_LOCAL_HMI_ACTIVE : BOOL;  (* DI 10016 | DIP1500 Local HMI Active *)
  SCADA_OUTPUT_FIRMWARE_VERSION : WORD;  (* IR 91 | DIP1500 Firmware Version | 3+5+8 bits (major+minor+revision) *)
  SCADA_OUTPUT_HARDWARE_VERSION : WORD;  (* IR 92 | DIP1500 Hardware Version | 3+5+8 bits (major+minor+revision) *)
  SCADA_OUTPUT_TEMPERATURE : WORD;  (* IR 93 | DIP1500 Temperature | degC | (raw - 500) / 10 *)
  SCADA_OUTPUT_FLOAT_LEVEL_ALARM : WORD;  (* IR 94 | DIP1500 Float Level Alarm *)
  SCADA_OUTPUT_DIGITAL_OUTPUT_VALUE : WORD;  (* IR 95 | DIP1500 Digital Output Value *)
  SCADA_OUTPUT_REAL_TIME_RUN_TIME_OR_VOLUME : DUT_Union_Real_Word;  (* IR 96-97 | DIP1500 Real-Time Run Time Or Volume | ms (time mode) / ml (volume mode) *)
  SCADA_OUTPUT_ACCUMULATED_RUN_TIME_OR_VOLUME : DUT_Union_Real_Word;  (* IR 98-99 | DIP1500 Accumulated Run Time Or Volume | ms (time mode) / ml (volume mode) *)
  HMI_INPUT_MOTOR_START_STOP : BOOL;  (* [HMI (local panel, FUXA address + 1000) : input (to PLC)] Coil 1003 | DIP1500 Motor Start Stop *)
  HMI_INPUT_MOTOR_DIRECTION : BOOL;  (* Coil 1004 | DIP1500 Motor Direction *)
  HMI_INPUT_FLASH_SAVE : BOOL;  (* Coil 1005 | DIP1500 Flash Save *)
  HMI_INPUT_OPERATION_MODE : BOOL;  (* Coil 1006 | DIP1500 Operation Mode *)
  HMI_INPUT_PARAM_WRITE_ENABLE : BOOL;  (* Coil 1007 | DIP1500 Parameter Write Enable *)
  HMI_INPUT_LOCAL_REQUEST : BOOL;  (* Coil 1010 | DIP1500 Local Request *)
  HMI_INPUT_AUTO_REQUEST : BOOL;  (* Coil 1011 | DIP1500 Auto Request *)
  HMI_INPUT_FOOT_SWITCH_INPUT_MODE : WORD;  (* HR 1009 | DIP1500 Foot Switch Input Mode *)
  HMI_INPUT_LIQUID_LEVEL_INPUT_MODE : WORD;  (* HR 1010 | DIP1500 Liquid Level Input Mode *)
  HMI_INPUT_STATE_OUTPUT_MODE : WORD;  (* HR 1011 | DIP1500 State Output Mode *)
  HMI_INPUT_COMMUNICATION_ADDRESS : WORD;  (* HR 1012 | DIP1500 Communication Address *)
  HMI_INPUT_BAUD_RATE_INDEX : WORD;  (* HR 1013 | DIP1500 Baud Rate Index | index *)
  HMI_INPUT_MOTOR_SPEED : DUT_Union_Real_Word;  (* HR 1001-1002 | DIP1500 Motor Speed | rpm *)
  HMI_INPUT_MAX_MOTOR_SPEED : DUT_Union_Real_Word;  (* HR 1003-1004 | DIP1500 Max Motor Speed | rpm *)
  HMI_INPUT_RUN_TIME_OR_VOLUME_SETPOINT : DUT_Union_Real_Word;  (* HR 1005-1006 | DIP1500 Run Time Or Volume Setpoint | ms (time mode) / ml (volume mode) *)
  HMI_INPUT_FLOW_RATE_OR_SPEED_CALIBRATION_COEFFICIENT : DUT_Union_Real_Word;  (* HR 1007-1008 | DIP1500 Flow Rate Or Speed Calibration Coefficient | ml/min or rpm *)
  HMI_OUTPUT_LOCAL_ACTIVE : BOOL;  (* [HMI (local panel, FUXA address + 1000) : output (from PLC)] DI 11016 | DIP1500 Local Active *)
  HMI_OUTPUT_FIRMWARE_VERSION : WORD;  (* IR 1091 | DIP1500 Firmware Version | 3+5+8 bits (major+minor+revision) *)
  HMI_OUTPUT_HARDWARE_VERSION : WORD;  (* IR 1092 | DIP1500 Hardware Version | 3+5+8 bits (major+minor+revision) *)
  HMI_OUTPUT_TEMPERATURE : WORD;  (* IR 1093 | DIP1500 Temperature | degC | (raw - 500) / 10 *)
  HMI_OUTPUT_FLOAT_LEVEL_ALARM : WORD;  (* IR 1094 | DIP1500 Float Level Alarm *)
  HMI_OUTPUT_DIGITAL_OUTPUT_VALUE : WORD;  (* IR 1095 | DIP1500 Digital Output Value *)
  HMI_OUTPUT_REAL_TIME_RUN_TIME_OR_VOLUME : DUT_Union_Real_Word;  (* IR 1096-1097 | DIP1500 Real-Time Run Time Or Volume | ms (time mode) / ml (volume mode) *)
  HMI_OUTPUT_ACCUMULATED_RUN_TIME_OR_VOLUME : DUT_Union_Real_Word;  (* IR 1098-1099 | DIP1500 Accumulated Run Time Or Volume | ms (time mode) / ml (volume mode) *)
  WEBVISU_INPUT_MOTOR_START_STOP : BOOL;  (* [WEBVISU : direct IEC variable] DIP1500 Motor Start Stop *)
  WEBVISU_INPUT_MOTOR_DIRECTION : BOOL;  (* [WEBVISU : direct IEC variable] DIP1500 Motor Direction *)
  WEBVISU_INPUT_FLASH_SAVE : BOOL;  (* [WEBVISU : direct IEC variable] DIP1500 Flash Save *)
  WEBVISU_INPUT_OPERATION_MODE : BOOL;  (* [WEBVISU : direct IEC variable] DIP1500 Operation Mode *)
  WEBVISU_INPUT_PARAM_WRITE_ENABLE : BOOL;  (* [WEBVISU : direct IEC variable] DIP1500 Parameter Write Enable *)
  WEBVISU_INPUT_LOCAL_REQUEST : BOOL;  (* [WEBVISU : direct IEC variable] DIP1500 Local Request *)
  WEBVISU_INPUT_AUTO_REQUEST : BOOL;  (* [WEBVISU : direct IEC variable] DIP1500 Auto Request *)
  WEBVISU_INPUT_FOOT_SWITCH_INPUT_MODE : WORD;  (* [WEBVISU : direct IEC variable] DIP1500 Foot Switch Input Mode *)
  WEBVISU_INPUT_LIQUID_LEVEL_INPUT_MODE : WORD;  (* [WEBVISU : direct IEC variable] DIP1500 Liquid Level Input Mode *)
  WEBVISU_INPUT_STATE_OUTPUT_MODE : WORD;  (* [WEBVISU : direct IEC variable] DIP1500 State Output Mode *)
  WEBVISU_INPUT_COMMUNICATION_ADDRESS : WORD;  (* [WEBVISU : direct IEC variable] DIP1500 Communication Address *)
  WEBVISU_INPUT_BAUD_RATE_INDEX : WORD;  (* [WEBVISU : direct IEC variable] DIP1500 Baud Rate Index | index *)
  WEBVISU_INPUT_MOTOR_SPEED : DUT_Union_Real_Word;  (* [WEBVISU : direct IEC variable] DIP1500 Motor Speed | rpm *)
  WEBVISU_INPUT_MAX_MOTOR_SPEED : DUT_Union_Real_Word;  (* [WEBVISU : direct IEC variable] DIP1500 Max Motor Speed | rpm *)
  WEBVISU_INPUT_RUN_TIME_OR_VOLUME_SETPOINT : DUT_Union_Real_Word;  (* [WEBVISU : direct IEC variable] DIP1500 Run Time Or Volume Setpoint | ms (time mode) / ml (volume mode) *)
  WEBVISU_INPUT_FLOW_RATE_OR_SPEED_CALIBRATION_COEFFICIENT : DUT_Union_Real_Word;  (* [WEBVISU : direct IEC variable] DIP1500 Flow Rate Or Speed Calibration Coefficient | ml/min or rpm *)
  WEBVISU_OUTPUT_LOCAL_ACTIVE : BOOL;  (* [WEBVISU : direct IEC variable] DIP1500 Local Active *)
  WEBVISU_OUTPUT_FIRMWARE_VERSION : WORD;  (* [WEBVISU : direct IEC variable] DIP1500 Firmware Version | 3+5+8 bits (major+minor+revision) *)
  WEBVISU_OUTPUT_HARDWARE_VERSION : WORD;  (* [WEBVISU : direct IEC variable] DIP1500 Hardware Version | 3+5+8 bits (major+minor+revision) *)
  WEBVISU_OUTPUT_TEMPERATURE : WORD;  (* [WEBVISU : direct IEC variable] DIP1500 Temperature | degC | (raw - 500) / 10 *)
  WEBVISU_OUTPUT_FLOAT_LEVEL_ALARM : WORD;  (* [WEBVISU : direct IEC variable] DIP1500 Float Level Alarm *)
  WEBVISU_OUTPUT_DIGITAL_OUTPUT_VALUE : WORD;  (* [WEBVISU : direct IEC variable] DIP1500 Digital Output Value *)
  WEBVISU_OUTPUT_REAL_TIME_RUN_TIME_OR_VOLUME : DUT_Union_Real_Word;  (* [WEBVISU : direct IEC variable] DIP1500 Real-Time Run Time Or Volume | ms (time mode) / ml (volume mode) *)
  WEBVISU_OUTPUT_ACCUMULATED_RUN_TIME_OR_VOLUME : DUT_Union_Real_Word;  (* [WEBVISU : direct IEC variable] DIP1500 Accumulated Run Time Or Volume | ms (time mode) / ml (volume mode) *)
  WEBVISU_OUTPUT_LOCAL_FUXA_ACTIVE : BOOL;  (* Effective FUXA local mode (masked by WEBVISU and HMI priority) *)
  WEBVISU_OUTPUT_LOCAL_HMI_ACTIVE : BOOL;  (* Effective HMI local mode (masked by WEBVISU priority) *)
END_STRUCT;
END_TYPE

TYPE DUT_EXC_DIP1500 : STRUCT
  UPI_INPUT_GLOBAL_LOCAL_FUXA : BOOL;  (* [UPI : functional units to equipment] From UPI_LOCAL_FUXA : global FUXA local active *)
  UPI_INPUT_GLOBAL_LOCAL_HMI : BOOL;  (* From UPI_LOCAL_HMI : global HMI local active *)
  UPI_INPUT_RUN : BOOL;  (* [UPI : commands used in auto mode] Auto mode command : run *)
  UPI_INPUT_CLOCKWISE : BOOL;  (* Auto mode command : 1 clockwise *)
  UPI_INPUT_VOLUME_MODE : BOOL;  (* Auto mode command : 0 time mode, 1 volume mode *)
  UPI_INPUT_SPEED : REAL;  (* Auto mode command : speed, rpm *)
  UPI_INPUT_RUN_SETPOINT : REAL;  (* Auto mode command : ms (time mode) or ml (volume mode), 0 = continuous *)
  UPI_INPUT_GLOBAL_LOCAL_WEBVISU : BOOL;  (* From UPI_LOCAL_WEBVISU : global WEBVISU local active *)
END_STRUCT;
END_TYPE

TYPE DUT_IO_DIP1500 : STRUCT
  SPARE : BOOL;  (* Placeholder, structure not used yet *)
END_STRUCT;
END_TYPE

TYPE DUT_PA_ADM100W : STRUCT
  SPARE : BOOL;  (* Placeholder, structure not used yet *)
END_STRUCT;
END_TYPE

TYPE DUT_PA_DOSENSOR : STRUCT
  SPARE : BOOL;  (* Placeholder, structure not used yet *)
END_STRUCT;
END_TYPE

TYPE DUT_COM_UPI_LOCAL_HMI : STRUCT
  SCADA_OUTPUT_LOCAL_ACTIVE : BOOL;  (* [SCADA (FUXA) : output (from PLC)] DI 10020 | Global Local HMI Active *)
  HMI_INPUT_LOCAL_REQUEST : BOOL;  (* [HMI (local panel, FUXA address + 1000) : input (to PLC)] Coil 1014 | Global Local HMI Request *)
  HMI_INPUT_AUTO_REQUEST : BOOL;  (* Coil 1015 | Global Auto HMI Request *)
  HMI_OUTPUT_LOCAL_ACTIVE : BOOL;  (* [HMI (local panel, FUXA address + 1000) : output (from PLC)] DI 11020 | Global Local HMI Active *)
END_STRUCT;
END_TYPE

TYPE DUT_EXC_UPI_LOCAL_FUXA : STRUCT
  UPI_OUTPUT_LOCAL_ACTIVE : BOOL;  (* [UPI : to equipment] Global FUXA local active *)
END_STRUCT;
END_TYPE

TYPE DUT_EXC_UPI_LOCAL_HMI : STRUCT
  UPI_OUTPUT_LOCAL_ACTIVE : BOOL;  (* [UPI : to equipment] Global HMI local active *)
END_STRUCT;
END_TYPE

TYPE DUT_INT_UPI_LOCAL_FUXA : STRUCT
  LOCAL_REQUEST : BOOL;  (* Local request (pulse or maintained) *)
  AUTO_REQUEST : BOOL;  (* Auto request, releases the global local *)
  LOCAL_ACTIVE : BOOL;  (* Memory : global local active *)
END_STRUCT;
END_TYPE

TYPE DUT_INT_UPI_LOCAL_HMI : STRUCT
  LOCAL_REQUEST : BOOL;  (* Local request (pulse or maintained) *)
  AUTO_REQUEST : BOOL;  (* Auto request, releases the global local *)
  LOCAL_ACTIVE : BOOL;  (* Memory : global local active *)
END_STRUCT;
END_TYPE

TYPE DUT_COM_UPI_LOCAL_WEBVISU : STRUCT
  WEBVISU_INPUT_LOCAL_REQUEST : BOOL;  (* [WEBVISU (direct IEC variables) : input (to PLC)] Global Local WEBVISU Request *)
  WEBVISU_INPUT_AUTO_REQUEST : BOOL;  (* Global Auto WEBVISU Request *)
  WEBVISU_OUTPUT_LOCAL_ACTIVE : BOOL;  (* [WEBVISU (direct IEC variables) : output (from PLC)] Global Local WEBVISU Active *)
END_STRUCT;
END_TYPE

TYPE DUT_EXC_UPI_LOCAL_WEBVISU : STRUCT
  UPI_OUTPUT_LOCAL_ACTIVE : BOOL;  (* [UPI : to equipment] Global WEBVISU local active *)
END_STRUCT;
END_TYPE

TYPE DUT_INT_UPI_LOCAL_WEBVISU : STRUCT
  LOCAL_REQUEST : BOOL;  (* Local request (pulse or maintained) *)
  AUTO_REQUEST : BOOL;  (* Auto request, releases the global local *)
  LOCAL_ACTIVE : BOOL;  (* Memory : global local active *)
END_STRUCT;
END_TYPE

TYPE DUT_INT_DIP1500 : STRUCT
  FUXA_LOCAL_REQUEST : BOOL;  (* [Control mode] From FUXA : local request (pulse or maintained) *)
  FUXA_AUTO_REQUEST : BOOL;  (* From FUXA : auto request, releases the individual FUXA local *)
  HMI_LOCAL_REQUEST : BOOL;  (* From HMI : local request (pulse or maintained) *)
  HMI_AUTO_REQUEST : BOOL;  (* From HMI : auto request, releases the individual HMI local *)
  GLOBAL_LOCAL_FUXA : BOOL;  (* From UPI_LOCAL_FUXA : global FUXA local active *)
  GLOBAL_LOCAL_HMI : BOOL;  (* From UPI_LOCAL_HMI : global HMI local active *)
  LOCAL_FUXA_INDIVIDUAL : BOOL;  (* Memory : individual FUXA local, set by local request, reset by auto request *)
  LOCAL_HMI_INDIVIDUAL : BOOL;  (* Memory : individual HMI local, set by local request, reset by auto request *)
  LOCAL_HMI : BOOL;  (* Result : equipment in HMI local (individual or global), unless WEBVISU local is active *)
  LOCAL_FUXA : BOOL;  (* Result : equipment in FUXA local (individual or global), unless WEBVISU or HMI local is active *)
  AUTO : BOOL;  (* Result : no local mode, commands come from the functional units (UPI) *)
  CMD_RUN : BOOL;  (* [Commands (to pump), from the active source] 0 stop, 1 start *)
  CMD_CLOCKWISE : BOOL;  (* 0 counterclockwise, 1 clockwise *)
  CMD_SAVE_FLASH : BOOL;  (* 1 s pulse to coil 0x0003, saves pump parameters to flash *)
  CMD_VOLUME_MODE : BOOL;  (* 0 time mode, 1 volume mode *)
  CMD_SPEED : REAL;  (* rpm *)
  CMD_MAX_SPEED : REAL;  (* rpm *)
  CMD_RUN_SETPOINT : REAL;  (* ms (time mode) or ml (volume mode), 0 = continuous *)
  CMD_CALIB_COEF : REAL;  (* ml/min or rpm *)
  CMD_FOOT_MODE : WORD;  (* Foot switch input mode *)
  CMD_LEVEL_MODE : WORD;  (* Liquid level input mode *)
  CMD_STATE_OUT_MODE : WORD;  (* State output mode *)
  CMD_ADDRESS : WORD;  (* Modbus address *)
  CMD_BAUD_INDEX : WORD;  (* 0=1200 .. 3=9600 .. 7=115200 *)
  PARAM_WRITE_ENABLE : BOOL;  (* [Parameter writing] 1 = write configuration to the pump, 0 = stop writing *)
  FLASH_SAVE_REQUEST : BOOL;  (* Flash save request (rising edge used) *)
  PARAM_VALID : BOOL;  (* Address 1..31, baud index 0..7, max speed > 0, calibration coefficient > 0 *)
  PULSE_500MS : BOOL;  (* [Write triggers] Square wave, 500 ms period, source of the trigger edges *)
  CMD_CHANGED : BOOL;  (* A command value changed this cycle *)
  CMD_WINDOW : BOOL;  (* Command write window, 3 s after the last change *)
  CMD_TRIGGER : BOOL;  (* Command channel trigger *)
  CONFIG_TRIGGER : BOOL;  (* Configuration channel trigger *)
  PREV_RUN : BOOL;  (* [Previous command values] Previous values for change detection *)
  PREV_CLOCKWISE : BOOL;
  PREV_VOLUME_MODE : BOOL;
  PREV_SAVE_FLASH : BOOL;
  PREV_SPEED : REAL;
  PREV_MAX_SPEED : REAL;
  PREV_RUN_SETPOINT : REAL;
  FBK_FIRMWARE_VERSION : WORD;  (* [Feedback (from pump)] 3+5+8 bits (major+minor+revision) *)
  FBK_HARDWARE_VERSION : WORD;  (* 3+5+8 bits (major+sub+reserved) *)
  FBK_TEMPERATURE : WORD;  (* (raw - 500) / 10 = degC, 65535 = not connected *)
  FBK_LEVEL_ALARM : WORD;  (* 0 no alarm, 1 alarm, 65535 = not connected *)
  FBK_DIGITAL_OUTPUT : WORD;  (* Digital output value *)
  FBK_RUN_ACTUAL : REAL;  (* Current run, ms (time mode) or ml (volume mode) *)
  FBK_RUN_TOTAL : REAL;  (* Accumulated run, ms (time mode) or ml (volume mode) *)
  UDINT_TEMP : UDINT;  (* [Work] Work variable, time mode conversion *)
  WEBVISU_LOCAL_REQUEST : BOOL;  (* From WEBVISU : individual local request *)
  WEBVISU_AUTO_REQUEST : BOOL;  (* From WEBVISU : releases individual WEBVISU local (auto wins) *)
  GLOBAL_LOCAL_WEBVISU : BOOL;  (* From UPI_LOCAL_WEBVISU : global local request *)
  LOCAL_WEBVISU_INDIVIDUAL : BOOL;  (* Memory : individual WEBVISU local request *)
  LOCAL_WEBVISU : BOOL;  (* Effective WEBVISU local : highest source priority *)
  SRC_MAX_MOTOR_SPEED : REAL;  (* [Parameter source] Value typed in the active local supervision *)
  SRC_CALIBRATION_COEFFICIENT : REAL;
  SRC_FOOT_SWITCH_INPUT_MODE : WORD;
  SRC_LIQUID_LEVEL_INPUT_MODE : WORD;
  SRC_STATE_OUTPUT_MODE : WORD;
  SRC_COMMUNICATION_ADDRESS : WORD;
  SRC_BAUD_RATE_INDEX : WORD;
  PREV_SRC_MAX_MOTOR_SPEED : REAL;  (* [Parameter change detection] Previous source values *)
  PREV_SRC_CALIBRATION_COEFFICIENT : REAL;
  PREV_SRC_FOOT_SWITCH_INPUT_MODE : WORD;
  PREV_SRC_LIQUID_LEVEL_INPUT_MODE : WORD;
  PREV_SRC_STATE_OUTPUT_MODE : WORD;
  PREV_SRC_COMMUNICATION_ADDRESS : WORD;
  PREV_SRC_BAUD_RATE_INDEX : WORD;
  PREV_LOCAL_WEBVISU : BOOL;  (* Previous control mode, to ignore the cycle where the source changes *)
  PREV_LOCAL_HMI : BOOL;
  PREV_LOCAL_FUXA : BOOL;
  SOURCE_CHANGED : BOOL;  (* The active local source changed this cycle : no parameter is taken *)
END_STRUCT;
END_TYPE

TYPE DUT_PA_DIP1500 : STRUCT
  MAX_MOTOR_SPEED : REAL := 350;  (* [Pump configuration, default value = declaration value, kept in GVL_PA (persistent)] rpm. Max motor speed (pump register 0x4003) *)
  CALIBRATION_COEFFICIENT : REAL := 100;  (* ml/min or rpm. Flow / speed calibration coefficient (0x400B) *)
  FOOT_SWITCH_INPUT_MODE : WORD := 0;  (* Foot switch input mode (0x400D) *)
  LIQUID_LEVEL_INPUT_MODE : WORD := 100;  (* Liquid level input mode (0x400E) *)
  STATE_OUTPUT_MODE : WORD := 7;  (* State output mode (0x400F) *)
  COMMUNICATION_ADDRESS : WORD := 11;  (* Pump Modbus address, 1..31 (0x4010) *)
  BAUD_RATE_INDEX : WORD := 3;  (* 0=1200 .. 3=9600 .. 7=115200 (0x4011) *)
END_STRUCT;
END_TYPE

VAR_GLOBAL  (* GVL_MODBUS *)
  Coils_TCP_HMI : ARRAY[0..187] OF BYTE;  (* -----------------Modbus TCP line IHM -> API (coils, %IX) *)
  Discret_input_TCP_HMI : ARRAY[0..187] OF BYTE;  (* API -> IHM (entrées discrètes, %QX) *)
  Holding_register_TCP_HMI : ARRAY[0..1500] OF WORD;  (* IHM -> API (registres de retenue, %IW) *)
  Input_register_TCP_HMI : ARRAY[0..1500] OF WORD;  (* API -> IHM (registres d'entrée, %QW) *)
  ADM100W_InputRegisters : ARRAY[0..87] OF WORD;  (* ------------------Modbus RTU line ---ADM100W *)
  ADM100W_Alarms : ARRAY[0..1] OF BYTE;
  DIP1500_Coils : ARRAY[0..3] OF BOOL;  (* ---Kamoer DIP1500 Coils - wrinting to pump *)
  DIP1500_InputRegisters : ARRAY[0..4] OF WORD;  (* input register - reading from pump *)
  DIP1500_Holding_Cmd : ARRAY[0..5] OF WORD;  (* Discrete input Holding registers - Writing to pump *)
  DIP1500_Holding_Config : ARRAY[0..6] OF WORD;
  DIP1500_Holding_Counters : ARRAY[0..3] OF WORD;  (* Holding registers - Reading from pump *)
END_VAR

{attribute 'qualified_only'}
VAR_GLOBAL  (* GVL_IO *)
  IO_ADM100W_1 : DUT_IO_ADM100W;  (* Trumeter ADM100W power meter *)
  IO_DOSENSOR_1 : DUT_IO_DOSENSOR;  (* Dissolved oxygen sensor *)
  IO_DIP1500_1 : DUT_IO_DIP1500;  (* Kamoer DIP1500 peristaltic pump *)
END_VAR

{attribute 'qualified_only'}
VAR_GLOBAL  (* GVL_IOMAP *)
  IOMAP_AI_SIGNAL_DOSENSOR_1 : DWORD;
  IOMAP_DI_FAULT_DOSENSOR_1 : BOOL;
  IOMAP_DO_HIGH_DOSENSOR_1 : BOOL;
  IOMAP_DO_LOW_DOSENSOR_1 : BOOL;
END_VAR

{attribute 'qualified_only'}
VAR_GLOBAL  (* GVL_COM *)
  COM_ADM100W_1 : DUT_COM_ADM100W;  (* Trumeter ADM100W power meter *)
  COM_DOSENSOR_1 : DUT_COM_DOSENSOR;  (* Dissolved oxygen sensor *)
  COM_DIP1500_1 : DUT_COM_DIP1500;  (* Kamoer DIP1500 peristaltic pump *)
  COM_UPI_LOCAL_FUXA : DUT_COM_UPI_LOCAL_FUXA;  (* Global FUXA local mode *)
  COM_UPI_LOCAL_HMI : DUT_COM_UPI_LOCAL_HMI;  (* Global HMI local mode *)
  COM_UPI_LOCAL_WEBVISU : DUT_COM_UPI_LOCAL_WEBVISU;  (* Global WEBVISU local mode *)
END_VAR

{attribute 'qualified_only'}
VAR_GLOBAL  (* GVL_EXC *)
  EXC_ADM100W_1 : DUT_EXC_ADM100W;  (* Trumeter ADM100W power meter *)
  EXC_DOSENSOR_1 : DUT_EXC_DOSENSOR;  (* Dissolved oxygen sensor *)
  EXC_DIP1500_1 : DUT_EXC_DIP1500;  (* Kamoer DIP1500 peristaltic pump *)
  EXC_UPI_LOCAL_FUXA : DUT_EXC_UPI_LOCAL_FUXA;  (* Global FUXA local mode *)
  EXC_UPI_LOCAL_HMI : DUT_EXC_UPI_LOCAL_HMI;  (* Global HMI local mode *)
  EXC_UPI_LOCAL_WEBVISU : DUT_EXC_UPI_LOCAL_WEBVISU;  (* Global WEBVISU local mode *)
END_VAR

{attribute 'qualified_only'}
{attribute 'checksumnoinit_override' := '3446479488'}
{attribute 'init_related_code' := '6eea8fa9-da21-468e-bab1-ddc04c20a5e9'}
VAR_GLOBAL RETAIN PERSISTENT  (* GVL_PA *)
  {attribute 'order_in_persistent_editor' := '0'}
  PA_ADM100W_1 : DUT_PA_ADM100W;  (* Trumeter ADM100W power meter *)
  {attribute 'order_in_persistent_editor' := '1'}
  PA_DOSENSOR_1 : DUT_PA_DOSENSOR;  (* Dissolved oxygen sensor *)
  {attribute 'order_in_persistent_editor' := '2'}
  PA_DIP1500_1 : DUT_PA_DIP1500;  (* Kamoer DIP1500 peristaltic pump *)
END_VAR

TYPE DUT_Union_Real_Word : UNION
  Real_value : REAL;
  Word_value : ARRAY[0..1] OF WORD;
END_UNION;
END_TYPE

PROGRAM PLC_PRG
  VAR
    GFB_UPI_1 : GFB_UPI;  (* Functional units *)
    GFB_INST_1 : GFB_INST;  (* Equipment instances *)
  END_VAR

            
//==============================================================================
// PLC_PRG
// Main cycle : 1. read all inputs, 2. functional units, 3. equipment, 4. write all outputs
//==============================================================================

//------------------------------------------------------------------------------
// 1. INPUTS : interfaces -> GVL
//------------------------------------------------------------------------------
GFC_COM_IN();
GFC_IO_IN();

//------------------------------------------------------------------------------
// 2. FUNCTIONAL UNITS (UPI) and their exchanges to the equipment
//------------------------------------------------------------------------------
GFB_UPI_1();
GFC_EXC_IN();

//------------------------------------------------------------------------------
// 3. EQUIPMENT
//------------------------------------------------------------------------------
GFB_INST_1();
GFC_EXC_OUT();

//------------------------------------------------------------------------------
// 4. OUTPUTS : GVL -> interfaces
//------------------------------------------------------------------------------
GFC_COM_OUT();
GFC_IO_OUT();

          
END_PROGRAM

FUNCTION FNC_REAL_TO_WORDS : BOOL
  VAR_INPUT
    Real_value : REAL;  (* Value to split *)
  END_VAR
  VAR_OUTPUT
    High_word : WORD;  (* Most significant word *)
    Low_word : WORD;  (* Least significant word *)
  END_VAR
  VAR
    Conversion : DUT_Union_Real_Word;  (* REAL / 2 WORD overlay *)
  END_VAR

            
//==============================================================================
// FNC_REAL_TO_WORDS
// REAL (IEEE 754) -> two Modbus words
// Call: FNC_REAL_TO_WORDS(Real_value := x, High_word => ..., Low_word => ...);
//==============================================================================

Conversion.Real_value := Real_value;
Low_word  := Conversion.Word_value[0];
High_word := Conversion.Word_value[1];
FNC_REAL_TO_WORDS := TRUE;

          
END_FUNCTION

FUNCTION FNC_WORDS_TO_REAL : REAL
  VAR_INPUT
    High_word : WORD;  (* Most significant word *)
    Low_word : WORD;  (* Least significant word *)
  END_VAR
  VAR
    Conversion : DUT_Union_Real_Word;  (* REAL / 2 WORD overlay *)
  END_VAR

            
//==============================================================================
// FNC_WORDS_TO_REAL
// Two Modbus words -> REAL (IEEE 754)
// ABCD device: High_word = lower address, CDAB device: Low_word = lower address
//==============================================================================

Conversion.Word_value[0] := Low_word;
Conversion.Word_value[1] := High_word;
FNC_WORDS_TO_REAL := Conversion.Real_value;

          
END_FUNCTION

FUNCTION GFC_COM_IN : BOOL

            
//==============================================================================
// GFC_COM_IN
// Modbus (GVL_MODBUS) -> GVL_COM : RTU equipment, SCADA FUXA, HMI
// Simple copies only, no conversion (conversions are done in the FBs)
//==============================================================================

//------------------------------------------------------------------------------
// COM : Modbus RTU, from equipment
//------------------------------------------------------------------------------
	//--- ADM100W_1
	GVL_COM.COM_ADM100W_1.COM_INPUT_IR    := GVL_MODBUS.ADM100W_InputRegisters;   // Input registers 0..87
	GVL_COM.COM_ADM100W_1.COM_INPUT_COILS := GVL_MODBUS.ADM100W_Alarms;           // Coils 0..9 (alarms)

	//--- DIP1500_1
	GVL_COM.COM_DIP1500_1.COM_INPUT_IR          := GVL_MODBUS.DIP1500_InputRegisters;     // Input registers 0x3001..0x3005
	GVL_COM.COM_DIP1500_1.COM_INPUT_HR_COUNTERS := GVL_MODBUS.DIP1500_Holding_Counters;   // Holding registers 0x4007..0x400A


//------------------------------------------------------------------------------
// SCADA FUXA : coils (FUXA 000001...)
//------------------------------------------------------------------------------
	//--- DOSENSOR_1
	GVL_COM.COM_DOSENSOR_1.SCADA_INPUT_CALIBRATION_HIGH := GVL_MODBUS.Coils_TCP_HMI[0].0;   // 1 | DO Calibration High
	GVL_COM.COM_DOSENSOR_1.SCADA_INPUT_CALIBRATION_LOW  := GVL_MODBUS.Coils_TCP_HMI[0].1;   // 2 | DO Calibration Low
	GVL_COM.COM_DOSENSOR_1.SCADA_INPUT_LOCAL_REQUEST    := GVL_MODBUS.Coils_TCP_HMI[0].7;   // 8 | DO Sensor Local Request
	GVL_COM.COM_DOSENSOR_1.SCADA_INPUT_AUTO_REQUEST     := GVL_MODBUS.Coils_TCP_HMI[1].0;   // 9 | DO Sensor Auto Request

	//--- DIP1500_1
	GVL_COM.COM_DIP1500_1.SCADA_INPUT_MOTOR_START_STOP   := GVL_MODBUS.Coils_TCP_HMI[0].2;   // 3 | DIP1500 Motor Start Stop
	GVL_COM.COM_DIP1500_1.SCADA_INPUT_MOTOR_DIRECTION    := GVL_MODBUS.Coils_TCP_HMI[0].3;   // 4 | DIP1500 Motor Direction
	GVL_COM.COM_DIP1500_1.SCADA_INPUT_FLASH_SAVE         := GVL_MODBUS.Coils_TCP_HMI[0].4;   // 5 | DIP1500 Flash Save
	GVL_COM.COM_DIP1500_1.SCADA_INPUT_OPERATION_MODE     := GVL_MODBUS.Coils_TCP_HMI[0].5;   // 6 | DIP1500 Operation Mode
	GVL_COM.COM_DIP1500_1.SCADA_INPUT_PARAM_WRITE_ENABLE := GVL_MODBUS.Coils_TCP_HMI[0].6;   // 7 | DIP1500 Parameter Write Enable
	GVL_COM.COM_DIP1500_1.SCADA_INPUT_LOCAL_REQUEST      := GVL_MODBUS.Coils_TCP_HMI[1].1;   // 10 | DIP1500 Local Request
	GVL_COM.COM_DIP1500_1.SCADA_INPUT_AUTO_REQUEST       := GVL_MODBUS.Coils_TCP_HMI[1].2;   // 11 | DIP1500 Auto Request

	//--- ADM100W_1
	GVL_COM.COM_ADM100W_1.SCADA_INPUT_LOCAL_REQUEST := GVL_MODBUS.Coils_TCP_HMI[1].3;   // 12 | ADM100W Local Request
	GVL_COM.COM_ADM100W_1.SCADA_INPUT_AUTO_REQUEST  := GVL_MODBUS.Coils_TCP_HMI[1].4;   // 13 | ADM100W Auto Request

	//--- UPI_LOCAL_FUXA
	GVL_COM.COM_UPI_LOCAL_FUXA.SCADA_INPUT_LOCAL_REQUEST := GVL_MODBUS.Coils_TCP_HMI[1].5;   // 14 | Global Local FUXA Request
	GVL_COM.COM_UPI_LOCAL_FUXA.SCADA_INPUT_AUTO_REQUEST  := GVL_MODBUS.Coils_TCP_HMI[1].6;   // 15 | Global Auto FUXA Request


//------------------------------------------------------------------------------
// SCADA FUXA : holding registers (FUXA 400001...), REAL = low word first (Float32MLE)
//------------------------------------------------------------------------------
	//--- DIP1500_1
	GVL_COM.COM_DIP1500_1.SCADA_INPUT_MOTOR_SPEED.Word_value[0]                                := GVL_MODBUS.Holding_register_TCP_HMI[0];    // 1 | DIP1500 Motor Speed (low word)
	GVL_COM.COM_DIP1500_1.SCADA_INPUT_MOTOR_SPEED.Word_value[1]                                := GVL_MODBUS.Holding_register_TCP_HMI[1];    // 2 | DIP1500 Motor Speed (high word)
	GVL_COM.COM_DIP1500_1.SCADA_INPUT_MAX_MOTOR_SPEED.Word_value[0]                            := GVL_MODBUS.Holding_register_TCP_HMI[2];    // 3 | DIP1500 Max Motor Speed (low word)
	GVL_COM.COM_DIP1500_1.SCADA_INPUT_MAX_MOTOR_SPEED.Word_value[1]                            := GVL_MODBUS.Holding_register_TCP_HMI[3];    // 4 | DIP1500 Max Motor Speed (high word)
	GVL_COM.COM_DIP1500_1.SCADA_INPUT_RUN_TIME_OR_VOLUME_SETPOINT.Word_value[0]                := GVL_MODBUS.Holding_register_TCP_HMI[4];    // 5 | DIP1500 Run Time Or Volume Setpoint (low word)
	GVL_COM.COM_DIP1500_1.SCADA_INPUT_RUN_TIME_OR_VOLUME_SETPOINT.Word_value[1]                := GVL_MODBUS.Holding_register_TCP_HMI[5];    // 6 | DIP1500 Run Time Or Volume Setpoint (high word)
	GVL_COM.COM_DIP1500_1.SCADA_INPUT_FLOW_RATE_OR_SPEED_CALIBRATION_COEFFICIENT.Word_value[0] := GVL_MODBUS.Holding_register_TCP_HMI[6];    // 7 | DIP1500 Flow Rate Or Speed Calibration Coefficient (low word)
	GVL_COM.COM_DIP1500_1.SCADA_INPUT_FLOW_RATE_OR_SPEED_CALIBRATION_COEFFICIENT.Word_value[1] := GVL_MODBUS.Holding_register_TCP_HMI[7];    // 8 | DIP1500 Flow Rate Or Speed Calibration Coefficient (high word)
	GVL_COM.COM_DIP1500_1.SCADA_INPUT_FOOT_SWITCH_INPUT_MODE                                   := GVL_MODBUS.Holding_register_TCP_HMI[8];    // 9 | DIP1500 Foot Switch Input Mode
	GVL_COM.COM_DIP1500_1.SCADA_INPUT_LIQUID_LEVEL_INPUT_MODE                                  := GVL_MODBUS.Holding_register_TCP_HMI[9];    // 10 | DIP1500 Liquid Level Input Mode
	GVL_COM.COM_DIP1500_1.SCADA_INPUT_STATE_OUTPUT_MODE                                        := GVL_MODBUS.Holding_register_TCP_HMI[10];   // 11 | DIP1500 State Output Mode
	GVL_COM.COM_DIP1500_1.SCADA_INPUT_COMMUNICATION_ADDRESS                                    := GVL_MODBUS.Holding_register_TCP_HMI[11];   // 12 | DIP1500 Communication Address
	GVL_COM.COM_DIP1500_1.SCADA_INPUT_BAUD_RATE_INDEX                                          := GVL_MODBUS.Holding_register_TCP_HMI[12];   // 13 | DIP1500 Baud Rate Index


//------------------------------------------------------------------------------
// HMI : coils (1001...)
//------------------------------------------------------------------------------
	//--- DOSENSOR_1
	GVL_COM.COM_DOSENSOR_1.HMI_INPUT_CALIBRATION_HIGH := GVL_MODBUS.Coils_TCP_HMI[125].0;   // 1001 | DO Calibration High
	GVL_COM.COM_DOSENSOR_1.HMI_INPUT_CALIBRATION_LOW  := GVL_MODBUS.Coils_TCP_HMI[125].1;   // 1002 | DO Calibration Low
	GVL_COM.COM_DOSENSOR_1.HMI_INPUT_LOCAL_REQUEST    := GVL_MODBUS.Coils_TCP_HMI[125].7;   // 1008 | DO Sensor Local Request
	GVL_COM.COM_DOSENSOR_1.HMI_INPUT_AUTO_REQUEST     := GVL_MODBUS.Coils_TCP_HMI[126].0;   // 1009 | DO Sensor Auto Request

	//--- DIP1500_1
	GVL_COM.COM_DIP1500_1.HMI_INPUT_MOTOR_START_STOP   := GVL_MODBUS.Coils_TCP_HMI[125].2;   // 1003 | DIP1500 Motor Start Stop
	GVL_COM.COM_DIP1500_1.HMI_INPUT_MOTOR_DIRECTION    := GVL_MODBUS.Coils_TCP_HMI[125].3;   // 1004 | DIP1500 Motor Direction
	GVL_COM.COM_DIP1500_1.HMI_INPUT_FLASH_SAVE         := GVL_MODBUS.Coils_TCP_HMI[125].4;   // 1005 | DIP1500 Flash Save
	GVL_COM.COM_DIP1500_1.HMI_INPUT_OPERATION_MODE     := GVL_MODBUS.Coils_TCP_HMI[125].5;   // 1006 | DIP1500 Operation Mode
	GVL_COM.COM_DIP1500_1.HMI_INPUT_PARAM_WRITE_ENABLE := GVL_MODBUS.Coils_TCP_HMI[125].6;   // 1007 | DIP1500 Parameter Write Enable
	GVL_COM.COM_DIP1500_1.HMI_INPUT_LOCAL_REQUEST      := GVL_MODBUS.Coils_TCP_HMI[126].1;   // 1010 | DIP1500 Local Request
	GVL_COM.COM_DIP1500_1.HMI_INPUT_AUTO_REQUEST       := GVL_MODBUS.Coils_TCP_HMI[126].2;   // 1011 | DIP1500 Auto Request

	//--- ADM100W_1
	GVL_COM.COM_ADM100W_1.HMI_INPUT_LOCAL_REQUEST := GVL_MODBUS.Coils_TCP_HMI[126].3;   // 1012 | ADM100W Local Request
	GVL_COM.COM_ADM100W_1.HMI_INPUT_AUTO_REQUEST  := GVL_MODBUS.Coils_TCP_HMI[126].4;   // 1013 | ADM100W Auto Request

	//--- UPI_LOCAL_HMI
	GVL_COM.COM_UPI_LOCAL_HMI.HMI_INPUT_LOCAL_REQUEST := GVL_MODBUS.Coils_TCP_HMI[126].5;   // 1014 | Global Local HMI Request
	GVL_COM.COM_UPI_LOCAL_HMI.HMI_INPUT_AUTO_REQUEST  := GVL_MODBUS.Coils_TCP_HMI[126].6;   // 1015 | Global Auto HMI Request


//------------------------------------------------------------------------------
// HMI : holding registers (1001...), REAL = low word first
//------------------------------------------------------------------------------
	//--- DIP1500_1
	GVL_COM.COM_DIP1500_1.HMI_INPUT_MOTOR_SPEED.Word_value[0]                                := GVL_MODBUS.Holding_register_TCP_HMI[1000];   // 1001 | DIP1500 Motor Speed (low word)
	GVL_COM.COM_DIP1500_1.HMI_INPUT_MOTOR_SPEED.Word_value[1]                                := GVL_MODBUS.Holding_register_TCP_HMI[1001];   // 1002 | DIP1500 Motor Speed (high word)
	GVL_COM.COM_DIP1500_1.HMI_INPUT_MAX_MOTOR_SPEED.Word_value[0]                            := GVL_MODBUS.Holding_register_TCP_HMI[1002];   // 1003 | DIP1500 Max Motor Speed (low word)
	GVL_COM.COM_DIP1500_1.HMI_INPUT_MAX_MOTOR_SPEED.Word_value[1]                            := GVL_MODBUS.Holding_register_TCP_HMI[1003];   // 1004 | DIP1500 Max Motor Speed (high word)
	GVL_COM.COM_DIP1500_1.HMI_INPUT_RUN_TIME_OR_VOLUME_SETPOINT.Word_value[0]                := GVL_MODBUS.Holding_register_TCP_HMI[1004];   // 1005 | DIP1500 Run Time Or Volume Setpoint (low word)
	GVL_COM.COM_DIP1500_1.HMI_INPUT_RUN_TIME_OR_VOLUME_SETPOINT.Word_value[1]                := GVL_MODBUS.Holding_register_TCP_HMI[1005];   // 1006 | DIP1500 Run Time Or Volume Setpoint (high word)
	GVL_COM.COM_DIP1500_1.HMI_INPUT_FLOW_RATE_OR_SPEED_CALIBRATION_COEFFICIENT.Word_value[0] := GVL_MODBUS.Holding_register_TCP_HMI[1006];   // 1007 | DIP1500 Flow Rate Or Speed Calibration Coefficient (low word)
	GVL_COM.COM_DIP1500_1.HMI_INPUT_FLOW_RATE_OR_SPEED_CALIBRATION_COEFFICIENT.Word_value[1] := GVL_MODBUS.Holding_register_TCP_HMI[1007];   // 1008 | DIP1500 Flow Rate Or Speed Calibration Coefficient (high word)
	GVL_COM.COM_DIP1500_1.HMI_INPUT_FOOT_SWITCH_INPUT_MODE                                   := GVL_MODBUS.Holding_register_TCP_HMI[1008];   // 1009 | DIP1500 Foot Switch Input Mode
	GVL_COM.COM_DIP1500_1.HMI_INPUT_LIQUID_LEVEL_INPUT_MODE                                  := GVL_MODBUS.Holding_register_TCP_HMI[1009];   // 1010 | DIP1500 Liquid Level Input Mode
	GVL_COM.COM_DIP1500_1.HMI_INPUT_STATE_OUTPUT_MODE                                        := GVL_MODBUS.Holding_register_TCP_HMI[1010];   // 1011 | DIP1500 State Output Mode
	GVL_COM.COM_DIP1500_1.HMI_INPUT_COMMUNICATION_ADDRESS                                    := GVL_MODBUS.Holding_register_TCP_HMI[1011];   // 1012 | DIP1500 Communication Address
	GVL_COM.COM_DIP1500_1.HMI_INPUT_BAUD_RATE_INDEX                                          := GVL_MODBUS.Holding_register_TCP_HMI[1012];   // 1013 | DIP1500 Baud Rate Index

GFC_COM_IN := TRUE;

          
END_FUNCTION

FUNCTION GFC_COM_OUT : BOOL

            
//==============================================================================
// GFC_COM_OUT
// GVL_COM -> Modbus (GVL_MODBUS) : RTU equipment, SCADA FUXA, HMI
// Simple copies only, no conversion (conversions are done in the FBs)
//==============================================================================

//------------------------------------------------------------------------------
// COM : Modbus RTU, to equipment (write triggers are mapped directly in the slave I/O mapping)
//------------------------------------------------------------------------------
	//--- DIP1500_1
	GVL_MODBUS.DIP1500_Coils          := GVL_COM.COM_DIP1500_1.COM_OUTPUT_COILS;       // Coils 0x0001..0x0004
	GVL_MODBUS.DIP1500_Holding_Cmd    := GVL_COM.COM_DIP1500_1.COM_OUTPUT_HR_CMD;      // Holding registers 0x4001..0x4006
	GVL_MODBUS.DIP1500_Holding_Config := GVL_COM.COM_DIP1500_1.COM_OUTPUT_HR_CONFIG;   // Holding registers 0x400B..0x4011


//------------------------------------------------------------------------------
// SCADA FUXA : discrete inputs (FUXA 100001...)
//------------------------------------------------------------------------------
	//--- DOSENSOR_1
	GVL_MODBUS.Discret_input_TCP_HMI[0].0 := GVL_COM.COM_DOSENSOR_1.SCADA_OUTPUT_FAULT;               // 10001 | Do sensor fault
	GVL_MODBUS.Discret_input_TCP_HMI[0].1 := GVL_COM.COM_DOSENSOR_1.SCADA_OUTPUT_CALIBRATION_DONE;    // 10002 | Do sensor calibration done
	GVL_MODBUS.Discret_input_TCP_HMI[1].4 := GVL_COM.COM_DOSENSOR_1.SCADA_OUTPUT_LOCAL_FUXA_ACTIVE;   // 10013 | DO Sensor Local FUXA Active
	GVL_MODBUS.Discret_input_TCP_HMI[1].5 := GVL_COM.COM_DOSENSOR_1.SCADA_OUTPUT_LOCAL_HMI_ACTIVE;    // 10014 | DO Sensor Local HMI Active

	//--- ADM100W_1
	GVL_MODBUS.Discret_input_TCP_HMI[0].2 := GVL_COM.COM_ADM100W_1.SCADA_OUTPUT_ALARM_1_STATUS;      // 10003 | ADM100W Alarm 1 Status
	GVL_MODBUS.Discret_input_TCP_HMI[0].3 := GVL_COM.COM_ADM100W_1.SCADA_OUTPUT_ALARM_2_STATUS;      // 10004 | ADM100W Alarm 2 Status
	GVL_MODBUS.Discret_input_TCP_HMI[0].4 := GVL_COM.COM_ADM100W_1.SCADA_OUTPUT_ALARM_3_STATUS;      // 10005 | ADM100W Alarm 3 Status
	GVL_MODBUS.Discret_input_TCP_HMI[0].5 := GVL_COM.COM_ADM100W_1.SCADA_OUTPUT_ALARM_4_STATUS;      // 10006 | ADM100W Alarm 4 Status
	GVL_MODBUS.Discret_input_TCP_HMI[0].6 := GVL_COM.COM_ADM100W_1.SCADA_OUTPUT_ALARM_5_STATUS;      // 10007 | ADM100W Alarm 5 Status
	GVL_MODBUS.Discret_input_TCP_HMI[0].7 := GVL_COM.COM_ADM100W_1.SCADA_OUTPUT_ALARM_6_STATUS;      // 10008 | ADM100W Alarm 6 Status
	GVL_MODBUS.Discret_input_TCP_HMI[1].0 := GVL_COM.COM_ADM100W_1.SCADA_OUTPUT_ALARM_7_STATUS;      // 10009 | ADM100W Alarm 7 Status
	GVL_MODBUS.Discret_input_TCP_HMI[1].1 := GVL_COM.COM_ADM100W_1.SCADA_OUTPUT_ALARM_8_STATUS;      // 10010 | ADM100W Alarm 8 Status
	GVL_MODBUS.Discret_input_TCP_HMI[1].2 := GVL_COM.COM_ADM100W_1.SCADA_OUTPUT_ALARM_9_STATUS;      // 10011 | ADM100W Alarm 9 Status
	GVL_MODBUS.Discret_input_TCP_HMI[1].3 := GVL_COM.COM_ADM100W_1.SCADA_OUTPUT_ALARM_10_STATUS;     // 10012 | ADM100W Alarm 10 Status
	GVL_MODBUS.Discret_input_TCP_HMI[2].0 := GVL_COM.COM_ADM100W_1.SCADA_OUTPUT_LOCAL_FUXA_ACTIVE;   // 10017 | ADM100W Local FUXA Active
	GVL_MODBUS.Discret_input_TCP_HMI[2].1 := GVL_COM.COM_ADM100W_1.SCADA_OUTPUT_LOCAL_HMI_ACTIVE;    // 10018 | ADM100W Local HMI Active

	//--- DIP1500_1
	GVL_MODBUS.Discret_input_TCP_HMI[1].6 := GVL_COM.COM_DIP1500_1.SCADA_OUTPUT_LOCAL_FUXA_ACTIVE;   // 10015 | DIP1500 Local FUXA Active
	GVL_MODBUS.Discret_input_TCP_HMI[1].7 := GVL_COM.COM_DIP1500_1.SCADA_OUTPUT_LOCAL_HMI_ACTIVE;    // 10016 | DIP1500 Local HMI Active

	//--- UPI_LOCAL_FUXA
	GVL_MODBUS.Discret_input_TCP_HMI[2].2 := GVL_COM.COM_UPI_LOCAL_FUXA.SCADA_OUTPUT_LOCAL_ACTIVE;   // 10019 | Global Local FUXA Active

	//--- UPI_LOCAL_HMI
	GVL_MODBUS.Discret_input_TCP_HMI[2].3 := GVL_COM.COM_UPI_LOCAL_HMI.SCADA_OUTPUT_LOCAL_ACTIVE;   // 10020 | Global Local HMI Active


//------------------------------------------------------------------------------
// SCADA FUXA : input registers (FUXA 300001...), REAL = low word first (Float32MLE)
//------------------------------------------------------------------------------
	//--- ADM100W_1
	GVL_MODBUS.Input_register_TCP_HMI[0]  := GVL_COM.COM_ADM100W_1.SCADA_OUTPUT_FREQUENCY.Word_value[0];                   // 1 | ADM100W Frequency (low word)
	GVL_MODBUS.Input_register_TCP_HMI[1]  := GVL_COM.COM_ADM100W_1.SCADA_OUTPUT_FREQUENCY.Word_value[1];                   // 2 | ADM100W Frequency (high word)
	GVL_MODBUS.Input_register_TCP_HMI[2]  := GVL_COM.COM_ADM100W_1.SCADA_OUTPUT_L1_L2_VOLTAGE.Word_value[0];               // 3 | ADM100W L1-L2 Voltage (low word)
	GVL_MODBUS.Input_register_TCP_HMI[3]  := GVL_COM.COM_ADM100W_1.SCADA_OUTPUT_L1_L2_VOLTAGE.Word_value[1];               // 4 | ADM100W L1-L2 Voltage (high word)
	GVL_MODBUS.Input_register_TCP_HMI[4]  := GVL_COM.COM_ADM100W_1.SCADA_OUTPUT_L1_N_VOLTAGE.Word_value[0];                // 5 | ADM100W L1-N Voltage (low word)
	GVL_MODBUS.Input_register_TCP_HMI[5]  := GVL_COM.COM_ADM100W_1.SCADA_OUTPUT_L1_N_VOLTAGE.Word_value[1];                // 6 | ADM100W L1-N Voltage (high word)
	GVL_MODBUS.Input_register_TCP_HMI[6]  := GVL_COM.COM_ADM100W_1.SCADA_OUTPUT_L1_CURRENT.Word_value[0];                  // 7 | ADM100W L1 Current (low word)
	GVL_MODBUS.Input_register_TCP_HMI[7]  := GVL_COM.COM_ADM100W_1.SCADA_OUTPUT_L1_CURRENT.Word_value[1];                  // 8 | ADM100W L1 Current (high word)
	GVL_MODBUS.Input_register_TCP_HMI[8]  := GVL_COM.COM_ADM100W_1.SCADA_OUTPUT_L1_ACTIVE_POWER.Word_value[0];             // 9 | ADM100W L1 Active Power (low word)
	GVL_MODBUS.Input_register_TCP_HMI[9]  := GVL_COM.COM_ADM100W_1.SCADA_OUTPUT_L1_ACTIVE_POWER.Word_value[1];             // 10 | ADM100W L1 Active Power (high word)
	GVL_MODBUS.Input_register_TCP_HMI[10] := GVL_COM.COM_ADM100W_1.SCADA_OUTPUT_L1_APPARENT_POWER.Word_value[0];           // 11 | ADM100W L1 Apparent Power (low word)
	GVL_MODBUS.Input_register_TCP_HMI[11] := GVL_COM.COM_ADM100W_1.SCADA_OUTPUT_L1_APPARENT_POWER.Word_value[1];           // 12 | ADM100W L1 Apparent Power (high word)
	GVL_MODBUS.Input_register_TCP_HMI[12] := GVL_COM.COM_ADM100W_1.SCADA_OUTPUT_L1_REACTIVE_POWER.Word_value[0];           // 13 | ADM100W L1 Reactive Power (low word)
	GVL_MODBUS.Input_register_TCP_HMI[13] := GVL_COM.COM_ADM100W_1.SCADA_OUTPUT_L1_REACTIVE_POWER.Word_value[1];           // 14 | ADM100W L1 Reactive Power (high word)
	GVL_MODBUS.Input_register_TCP_HMI[14] := GVL_COM.COM_ADM100W_1.SCADA_OUTPUT_L1_CURRENT_PHASE_ANGLE.Word_value[0];      // 15 | ADM100W L1 Current Phase Angle (low word)
	GVL_MODBUS.Input_register_TCP_HMI[15] := GVL_COM.COM_ADM100W_1.SCADA_OUTPUT_L1_CURRENT_PHASE_ANGLE.Word_value[1];      // 16 | ADM100W L1 Current Phase Angle (high word)
	GVL_MODBUS.Input_register_TCP_HMI[16] := GVL_COM.COM_ADM100W_1.SCADA_OUTPUT_L1_POWER_FACTOR.Word_value[0];             // 17 | ADM100W L1 Power Factor (low word)
	GVL_MODBUS.Input_register_TCP_HMI[17] := GVL_COM.COM_ADM100W_1.SCADA_OUTPUT_L1_POWER_FACTOR.Word_value[1];             // 18 | ADM100W L1 Power Factor (high word)
	GVL_MODBUS.Input_register_TCP_HMI[18] := GVL_COM.COM_ADM100W_1.SCADA_OUTPUT_L1_VOLTAGE_THD.Word_value[0];              // 19 | ADM100W L1 Voltage THD (low word)
	GVL_MODBUS.Input_register_TCP_HMI[19] := GVL_COM.COM_ADM100W_1.SCADA_OUTPUT_L1_VOLTAGE_THD.Word_value[1];              // 20 | ADM100W L1 Voltage THD (high word)
	GVL_MODBUS.Input_register_TCP_HMI[20] := GVL_COM.COM_ADM100W_1.SCADA_OUTPUT_L1_CURRENT_THD.Word_value[0];              // 21 | ADM100W L1 Current THD (low word)
	GVL_MODBUS.Input_register_TCP_HMI[21] := GVL_COM.COM_ADM100W_1.SCADA_OUTPUT_L1_CURRENT_THD.Word_value[1];              // 22 | ADM100W L1 Current THD (high word)
	GVL_MODBUS.Input_register_TCP_HMI[22] := GVL_COM.COM_ADM100W_1.SCADA_OUTPUT_L1_MAX_LOAD.Word_value[0];                 // 23 | ADM100W L1 Max Load (low word)
	GVL_MODBUS.Input_register_TCP_HMI[23] := GVL_COM.COM_ADM100W_1.SCADA_OUTPUT_L1_MAX_LOAD.Word_value[1];                 // 24 | ADM100W L1 Max Load (high word)
	GVL_MODBUS.Input_register_TCP_HMI[24] := GVL_COM.COM_ADM100W_1.SCADA_OUTPUT_L1_L2_VOLTAGE_PHASE_ANGLE.Word_value[0];   // 25 | ADM100W L1-L2 Voltage Phase Angle (low word)
	GVL_MODBUS.Input_register_TCP_HMI[25] := GVL_COM.COM_ADM100W_1.SCADA_OUTPUT_L1_L2_VOLTAGE_PHASE_ANGLE.Word_value[1];   // 26 | ADM100W L1-L2 Voltage Phase Angle (high word)
	GVL_MODBUS.Input_register_TCP_HMI[26] := GVL_COM.COM_ADM100W_1.SCADA_OUTPUT_L2_L3_VOLTAGE.Word_value[0];               // 27 | ADM100W L2-L3 Voltage (low word)
	GVL_MODBUS.Input_register_TCP_HMI[27] := GVL_COM.COM_ADM100W_1.SCADA_OUTPUT_L2_L3_VOLTAGE.Word_value[1];               // 28 | ADM100W L2-L3 Voltage (high word)
	GVL_MODBUS.Input_register_TCP_HMI[28] := GVL_COM.COM_ADM100W_1.SCADA_OUTPUT_L2_N_VOLTAGE.Word_value[0];                // 29 | ADM100W L2-N Voltage (low word)
	GVL_MODBUS.Input_register_TCP_HMI[29] := GVL_COM.COM_ADM100W_1.SCADA_OUTPUT_L2_N_VOLTAGE.Word_value[1];                // 30 | ADM100W L2-N Voltage (high word)
	GVL_MODBUS.Input_register_TCP_HMI[30] := GVL_COM.COM_ADM100W_1.SCADA_OUTPUT_L2_CURRENT.Word_value[0];                  // 31 | ADM100W L2 Current (low word)
	GVL_MODBUS.Input_register_TCP_HMI[31] := GVL_COM.COM_ADM100W_1.SCADA_OUTPUT_L2_CURRENT.Word_value[1];                  // 32 | ADM100W L2 Current (high word)
	GVL_MODBUS.Input_register_TCP_HMI[32] := GVL_COM.COM_ADM100W_1.SCADA_OUTPUT_L2_ACTIVE_POWER.Word_value[0];             // 33 | ADM100W L2 Active Power (low word)
	GVL_MODBUS.Input_register_TCP_HMI[33] := GVL_COM.COM_ADM100W_1.SCADA_OUTPUT_L2_ACTIVE_POWER.Word_value[1];             // 34 | ADM100W L2 Active Power (high word)
	GVL_MODBUS.Input_register_TCP_HMI[34] := GVL_COM.COM_ADM100W_1.SCADA_OUTPUT_L2_APPARENT_POWER.Word_value[0];           // 35 | ADM100W L2 Apparent Power (low word)
	GVL_MODBUS.Input_register_TCP_HMI[35] := GVL_COM.COM_ADM100W_1.SCADA_OUTPUT_L2_APPARENT_POWER.Word_value[1];           // 36 | ADM100W L2 Apparent Power (high word)
	GVL_MODBUS.Input_register_TCP_HMI[36] := GVL_COM.COM_ADM100W_1.SCADA_OUTPUT_L2_REACTIVE_POWER.Word_value[0];           // 37 | ADM100W L2 Reactive Power (low word)
	GVL_MODBUS.Input_register_TCP_HMI[37] := GVL_COM.COM_ADM100W_1.SCADA_OUTPUT_L2_REACTIVE_POWER.Word_value[1];           // 38 | ADM100W L2 Reactive Power (high word)
	GVL_MODBUS.Input_register_TCP_HMI[38] := GVL_COM.COM_ADM100W_1.SCADA_OUTPUT_L2_CURRENT_PHASE_ANGLE.Word_value[0];      // 39 | ADM100W L2 Current Phase Angle (low word)
	GVL_MODBUS.Input_register_TCP_HMI[39] := GVL_COM.COM_ADM100W_1.SCADA_OUTPUT_L2_CURRENT_PHASE_ANGLE.Word_value[1];      // 40 | ADM100W L2 Current Phase Angle (high word)
	GVL_MODBUS.Input_register_TCP_HMI[40] := GVL_COM.COM_ADM100W_1.SCADA_OUTPUT_L2_POWER_FACTOR.Word_value[0];             // 41 | ADM100W L2 Power Factor (low word)
	GVL_MODBUS.Input_register_TCP_HMI[41] := GVL_COM.COM_ADM100W_1.SCADA_OUTPUT_L2_POWER_FACTOR.Word_value[1];             // 42 | ADM100W L2 Power Factor (high word)
	GVL_MODBUS.Input_register_TCP_HMI[42] := GVL_COM.COM_ADM100W_1.SCADA_OUTPUT_L2_VOLTAGE_THD.Word_value[0];              // 43 | ADM100W L2 Voltage THD (low word)
	GVL_MODBUS.Input_register_TCP_HMI[43] := GVL_COM.COM_ADM100W_1.SCADA_OUTPUT_L2_VOLTAGE_THD.Word_value[1];              // 44 | ADM100W L2 Voltage THD (high word)
	GVL_MODBUS.Input_register_TCP_HMI[44] := GVL_COM.COM_ADM100W_1.SCADA_OUTPUT_L2_CURRENT_THD.Word_value[0];              // 45 | ADM100W L2 Current THD (low word)
	GVL_MODBUS.Input_register_TCP_HMI[45] := GVL_COM.COM_ADM100W_1.SCADA_OUTPUT_L2_CURRENT_THD.Word_value[1];              // 46 | ADM100W L2 Current THD (high word)
	GVL_MODBUS.Input_register_TCP_HMI[46] := GVL_COM.COM_ADM100W_1.SCADA_OUTPUT_L2_MAX_LOAD.Word_value[0];                 // 47 | ADM100W L2 Max Load (low word)
	GVL_MODBUS.Input_register_TCP_HMI[47] := GVL_COM.COM_ADM100W_1.SCADA_OUTPUT_L2_MAX_LOAD.Word_value[1];                 // 48 | ADM100W L2 Max Load (high word)
	GVL_MODBUS.Input_register_TCP_HMI[48] := GVL_COM.COM_ADM100W_1.SCADA_OUTPUT_L1_L3_VOLTAGE_PHASE_ANGLE.Word_value[0];   // 49 | ADM100W L1-L3 Voltage Phase Angle (low word)
	GVL_MODBUS.Input_register_TCP_HMI[49] := GVL_COM.COM_ADM100W_1.SCADA_OUTPUT_L1_L3_VOLTAGE_PHASE_ANGLE.Word_value[1];   // 50 | ADM100W L1-L3 Voltage Phase Angle (high word)
	GVL_MODBUS.Input_register_TCP_HMI[50] := GVL_COM.COM_ADM100W_1.SCADA_OUTPUT_L3_L1_VOLTAGE.Word_value[0];               // 51 | ADM100W L3-L1 Voltage (low word)
	GVL_MODBUS.Input_register_TCP_HMI[51] := GVL_COM.COM_ADM100W_1.SCADA_OUTPUT_L3_L1_VOLTAGE.Word_value[1];               // 52 | ADM100W L3-L1 Voltage (high word)
	GVL_MODBUS.Input_register_TCP_HMI[52] := GVL_COM.COM_ADM100W_1.SCADA_OUTPUT_L3_N_VOLTAGE.Word_value[0];                // 53 | ADM100W L3-N Voltage (low word)
	GVL_MODBUS.Input_register_TCP_HMI[53] := GVL_COM.COM_ADM100W_1.SCADA_OUTPUT_L3_N_VOLTAGE.Word_value[1];                // 54 | ADM100W L3-N Voltage (high word)
	GVL_MODBUS.Input_register_TCP_HMI[54] := GVL_COM.COM_ADM100W_1.SCADA_OUTPUT_L3_CURRENT.Word_value[0];                  // 55 | ADM100W L3 Current (low word)
	GVL_MODBUS.Input_register_TCP_HMI[55] := GVL_COM.COM_ADM100W_1.SCADA_OUTPUT_L3_CURRENT.Word_value[1];                  // 56 | ADM100W L3 Current (high word)
	GVL_MODBUS.Input_register_TCP_HMI[56] := GVL_COM.COM_ADM100W_1.SCADA_OUTPUT_L3_ACTIVE_POWER.Word_value[0];             // 57 | ADM100W L3 Active Power (low word)
	GVL_MODBUS.Input_register_TCP_HMI[57] := GVL_COM.COM_ADM100W_1.SCADA_OUTPUT_L3_ACTIVE_POWER.Word_value[1];             // 58 | ADM100W L3 Active Power (high word)
	GVL_MODBUS.Input_register_TCP_HMI[58] := GVL_COM.COM_ADM100W_1.SCADA_OUTPUT_L3_APPARENT_POWER.Word_value[0];           // 59 | ADM100W L3 Apparent Power (low word)
	GVL_MODBUS.Input_register_TCP_HMI[59] := GVL_COM.COM_ADM100W_1.SCADA_OUTPUT_L3_APPARENT_POWER.Word_value[1];           // 60 | ADM100W L3 Apparent Power (high word)
	GVL_MODBUS.Input_register_TCP_HMI[60] := GVL_COM.COM_ADM100W_1.SCADA_OUTPUT_L3_REACTIVE_POWER.Word_value[0];           // 61 | ADM100W L3 Reactive Power (low word)
	GVL_MODBUS.Input_register_TCP_HMI[61] := GVL_COM.COM_ADM100W_1.SCADA_OUTPUT_L3_REACTIVE_POWER.Word_value[1];           // 62 | ADM100W L3 Reactive Power (high word)
	GVL_MODBUS.Input_register_TCP_HMI[62] := GVL_COM.COM_ADM100W_1.SCADA_OUTPUT_L3_CURRENT_PHASE_ANGLE.Word_value[0];      // 63 | ADM100W L3 Current Phase Angle (low word)
	GVL_MODBUS.Input_register_TCP_HMI[63] := GVL_COM.COM_ADM100W_1.SCADA_OUTPUT_L3_CURRENT_PHASE_ANGLE.Word_value[1];      // 64 | ADM100W L3 Current Phase Angle (high word)
	GVL_MODBUS.Input_register_TCP_HMI[64] := GVL_COM.COM_ADM100W_1.SCADA_OUTPUT_L3_POWER_FACTOR.Word_value[0];             // 65 | ADM100W L3 Power Factor (low word)
	GVL_MODBUS.Input_register_TCP_HMI[65] := GVL_COM.COM_ADM100W_1.SCADA_OUTPUT_L3_POWER_FACTOR.Word_value[1];             // 66 | ADM100W L3 Power Factor (high word)
	GVL_MODBUS.Input_register_TCP_HMI[66] := GVL_COM.COM_ADM100W_1.SCADA_OUTPUT_L3_VOLTAGE_THD.Word_value[0];              // 67 | ADM100W L3 Voltage THD (low word)
	GVL_MODBUS.Input_register_TCP_HMI[67] := GVL_COM.COM_ADM100W_1.SCADA_OUTPUT_L3_VOLTAGE_THD.Word_value[1];              // 68 | ADM100W L3 Voltage THD (high word)
	GVL_MODBUS.Input_register_TCP_HMI[68] := GVL_COM.COM_ADM100W_1.SCADA_OUTPUT_L3_CURRENT_THD.Word_value[0];              // 69 | ADM100W L3 Current THD (low word)
	GVL_MODBUS.Input_register_TCP_HMI[69] := GVL_COM.COM_ADM100W_1.SCADA_OUTPUT_L3_CURRENT_THD.Word_value[1];              // 70 | ADM100W L3 Current THD (high word)
	GVL_MODBUS.Input_register_TCP_HMI[70] := GVL_COM.COM_ADM100W_1.SCADA_OUTPUT_L3_MAX_LOAD.Word_value[0];                 // 71 | ADM100W L3 Max Load (low word)
	GVL_MODBUS.Input_register_TCP_HMI[71] := GVL_COM.COM_ADM100W_1.SCADA_OUTPUT_L3_MAX_LOAD.Word_value[1];                 // 72 | ADM100W L3 Max Load (high word)
	GVL_MODBUS.Input_register_TCP_HMI[72] := GVL_COM.COM_ADM100W_1.SCADA_OUTPUT_INTERNAL_TEMPERATURE.Word_value[0];        // 73 | ADM100W Internal Temperature (low word)
	GVL_MODBUS.Input_register_TCP_HMI[73] := GVL_COM.COM_ADM100W_1.SCADA_OUTPUT_INTERNAL_TEMPERATURE.Word_value[1];        // 74 | ADM100W Internal Temperature (high word)
	GVL_MODBUS.Input_register_TCP_HMI[74] := GVL_COM.COM_ADM100W_1.SCADA_OUTPUT_ACTIVE_ENERGY.Word_value[0];               // 75 | ADM100W Active Energy (low word)
	GVL_MODBUS.Input_register_TCP_HMI[75] := GVL_COM.COM_ADM100W_1.SCADA_OUTPUT_ACTIVE_ENERGY.Word_value[1];               // 76 | ADM100W Active Energy (high word)
	GVL_MODBUS.Input_register_TCP_HMI[76] := GVL_COM.COM_ADM100W_1.SCADA_OUTPUT_APPARENT_ENERGY.Word_value[0];             // 77 | ADM100W Apparent Energy (low word)
	GVL_MODBUS.Input_register_TCP_HMI[77] := GVL_COM.COM_ADM100W_1.SCADA_OUTPUT_APPARENT_ENERGY.Word_value[1];             // 78 | ADM100W Apparent Energy (high word)
	GVL_MODBUS.Input_register_TCP_HMI[78] := GVL_COM.COM_ADM100W_1.SCADA_OUTPUT_REACTIVE_ENERGY.Word_value[0];             // 79 | ADM100W Reactive Energy (low word)
	GVL_MODBUS.Input_register_TCP_HMI[79] := GVL_COM.COM_ADM100W_1.SCADA_OUTPUT_REACTIVE_ENERGY.Word_value[1];             // 80 | ADM100W Reactive Energy (high word)
	GVL_MODBUS.Input_register_TCP_HMI[80] := GVL_COM.COM_ADM100W_1.SCADA_OUTPUT_TOTAL_ACTIVE_POWER.Word_value[0];          // 81 | ADM100W Total Active Power (low word)
	GVL_MODBUS.Input_register_TCP_HMI[81] := GVL_COM.COM_ADM100W_1.SCADA_OUTPUT_TOTAL_ACTIVE_POWER.Word_value[1];          // 82 | ADM100W Total Active Power (high word)
	GVL_MODBUS.Input_register_TCP_HMI[82] := GVL_COM.COM_ADM100W_1.SCADA_OUTPUT_TOTAL_APPARENT_POWER.Word_value[0];        // 83 | ADM100W Total Apparent Power (low word)
	GVL_MODBUS.Input_register_TCP_HMI[83] := GVL_COM.COM_ADM100W_1.SCADA_OUTPUT_TOTAL_APPARENT_POWER.Word_value[1];        // 84 | ADM100W Total Apparent Power (high word)
	GVL_MODBUS.Input_register_TCP_HMI[84] := GVL_COM.COM_ADM100W_1.SCADA_OUTPUT_TOTAL_REACTIVE_POWER.Word_value[0];        // 85 | ADM100W Total Reactive Power (low word)
	GVL_MODBUS.Input_register_TCP_HMI[85] := GVL_COM.COM_ADM100W_1.SCADA_OUTPUT_TOTAL_REACTIVE_POWER.Word_value[1];        // 86 | ADM100W Total Reactive Power (high word)
	GVL_MODBUS.Input_register_TCP_HMI[86] := GVL_COM.COM_ADM100W_1.SCADA_OUTPUT_ALL_PHASE_POWER_FACTOR.Word_value[0];      // 87 | ADM100W All Phase Power Factor (low word)
	GVL_MODBUS.Input_register_TCP_HMI[87] := GVL_COM.COM_ADM100W_1.SCADA_OUTPUT_ALL_PHASE_POWER_FACTOR.Word_value[1];      // 88 | ADM100W All Phase Power Factor (high word)

	//--- DOSENSOR_1
	GVL_MODBUS.Input_register_TCP_HMI[88] := GVL_COM.COM_DOSENSOR_1.SCADA_OUTPUT_SIGNAL.Word_value[0];   // 89 | DO Sensor Signal (low word)
	GVL_MODBUS.Input_register_TCP_HMI[89] := GVL_COM.COM_DOSENSOR_1.SCADA_OUTPUT_SIGNAL.Word_value[1];   // 90 | DO Sensor Signal (high word)

	//--- DIP1500_1
	GVL_MODBUS.Input_register_TCP_HMI[90] := GVL_COM.COM_DIP1500_1.SCADA_OUTPUT_FIRMWARE_VERSION;                               // 91 | DIP1500 Firmware Version
	GVL_MODBUS.Input_register_TCP_HMI[91] := GVL_COM.COM_DIP1500_1.SCADA_OUTPUT_HARDWARE_VERSION;                               // 92 | DIP1500 Hardware Version
	GVL_MODBUS.Input_register_TCP_HMI[92] := GVL_COM.COM_DIP1500_1.SCADA_OUTPUT_TEMPERATURE;                                    // 93 | DIP1500 Temperature
	GVL_MODBUS.Input_register_TCP_HMI[93] := GVL_COM.COM_DIP1500_1.SCADA_OUTPUT_FLOAT_LEVEL_ALARM;                              // 94 | DIP1500 Float Level Alarm
	GVL_MODBUS.Input_register_TCP_HMI[94] := GVL_COM.COM_DIP1500_1.SCADA_OUTPUT_DIGITAL_OUTPUT_VALUE;                           // 95 | DIP1500 Digital Output Value
	GVL_MODBUS.Input_register_TCP_HMI[95] := GVL_COM.COM_DIP1500_1.SCADA_OUTPUT_REAL_TIME_RUN_TIME_OR_VOLUME.Word_value[0];     // 96 | DIP1500 Real-Time Run Time Or Volume (low word)
	GVL_MODBUS.Input_register_TCP_HMI[96] := GVL_COM.COM_DIP1500_1.SCADA_OUTPUT_REAL_TIME_RUN_TIME_OR_VOLUME.Word_value[1];     // 97 | DIP1500 Real-Time Run Time Or Volume (high word)
	GVL_MODBUS.Input_register_TCP_HMI[97] := GVL_COM.COM_DIP1500_1.SCADA_OUTPUT_ACCUMULATED_RUN_TIME_OR_VOLUME.Word_value[0];   // 98 | DIP1500 Accumulated Run Time Or Volume (low word)
	GVL_MODBUS.Input_register_TCP_HMI[98] := GVL_COM.COM_DIP1500_1.SCADA_OUTPUT_ACCUMULATED_RUN_TIME_OR_VOLUME.Word_value[1];   // 99 | DIP1500 Accumulated Run Time Or Volume (high word)


//------------------------------------------------------------------------------
// HMI : discrete inputs (11001...)
//------------------------------------------------------------------------------
	//--- DOSENSOR_1
	GVL_MODBUS.Discret_input_TCP_HMI[125].0 := GVL_COM.COM_DOSENSOR_1.HMI_OUTPUT_FAULT;              // 11001 | Do sensor fault
	GVL_MODBUS.Discret_input_TCP_HMI[125].1 := GVL_COM.COM_DOSENSOR_1.HMI_OUTPUT_CALIBRATION_DONE;   // 11002 | Do sensor calibration done
	GVL_MODBUS.Discret_input_TCP_HMI[126].5 := GVL_COM.COM_DOSENSOR_1.HMI_OUTPUT_LOCAL_ACTIVE;       // 11014 | DO Sensor Local Active

	//--- ADM100W_1
	GVL_MODBUS.Discret_input_TCP_HMI[125].2 := GVL_COM.COM_ADM100W_1.HMI_OUTPUT_ALARM_1_STATUS;    // 11003 | ADM100W Alarm 1 Status
	GVL_MODBUS.Discret_input_TCP_HMI[125].3 := GVL_COM.COM_ADM100W_1.HMI_OUTPUT_ALARM_2_STATUS;    // 11004 | ADM100W Alarm 2 Status
	GVL_MODBUS.Discret_input_TCP_HMI[125].4 := GVL_COM.COM_ADM100W_1.HMI_OUTPUT_ALARM_3_STATUS;    // 11005 | ADM100W Alarm 3 Status
	GVL_MODBUS.Discret_input_TCP_HMI[125].5 := GVL_COM.COM_ADM100W_1.HMI_OUTPUT_ALARM_4_STATUS;    // 11006 | ADM100W Alarm 4 Status
	GVL_MODBUS.Discret_input_TCP_HMI[125].6 := GVL_COM.COM_ADM100W_1.HMI_OUTPUT_ALARM_5_STATUS;    // 11007 | ADM100W Alarm 5 Status
	GVL_MODBUS.Discret_input_TCP_HMI[125].7 := GVL_COM.COM_ADM100W_1.HMI_OUTPUT_ALARM_6_STATUS;    // 11008 | ADM100W Alarm 6 Status
	GVL_MODBUS.Discret_input_TCP_HMI[126].0 := GVL_COM.COM_ADM100W_1.HMI_OUTPUT_ALARM_7_STATUS;    // 11009 | ADM100W Alarm 7 Status
	GVL_MODBUS.Discret_input_TCP_HMI[126].1 := GVL_COM.COM_ADM100W_1.HMI_OUTPUT_ALARM_8_STATUS;    // 11010 | ADM100W Alarm 8 Status
	GVL_MODBUS.Discret_input_TCP_HMI[126].2 := GVL_COM.COM_ADM100W_1.HMI_OUTPUT_ALARM_9_STATUS;    // 11011 | ADM100W Alarm 9 Status
	GVL_MODBUS.Discret_input_TCP_HMI[126].3 := GVL_COM.COM_ADM100W_1.HMI_OUTPUT_ALARM_10_STATUS;   // 11012 | ADM100W Alarm 10 Status
	GVL_MODBUS.Discret_input_TCP_HMI[127].1 := GVL_COM.COM_ADM100W_1.HMI_OUTPUT_LOCAL_ACTIVE;      // 11018 | ADM100W Local Active

	//--- DIP1500_1
	GVL_MODBUS.Discret_input_TCP_HMI[126].7 := GVL_COM.COM_DIP1500_1.HMI_OUTPUT_LOCAL_ACTIVE;   // 11016 | DIP1500 Local Active

	//--- UPI_LOCAL_HMI
	GVL_MODBUS.Discret_input_TCP_HMI[127].3 := GVL_COM.COM_UPI_LOCAL_HMI.HMI_OUTPUT_LOCAL_ACTIVE;   // 11020 | Global Local HMI Active


